{region 'Documentation'}
(*!
<summary>Contributes only the checking Assertions, not the intentionally controlled subject results.</summary>
*)
{endregion}
METHOD PROTECTED AggregateResults
VAR_INPUT
    Aggregator : I_ResultAggregator; //! Borrowed result sink owned by the outer Test Case; add this test's checking Assertions without resetting or retaining the sink.
END_VAR
Aggregator.AddProvider(Provider := FInitialization);
Aggregator.AddProvider(Provider := FConfigureOrder);
Aggregator.AddProvider(Provider := FCollection);
Aggregator.AddProvider(Provider := FPassiveState);
Aggregator.AddProvider(Provider := FDiagnostic);
Aggregator.AddProvider(Provider := FDispatch);
Aggregator.AddProvider(Provider := FCaptureIntegrity);
END_METHOD

{region 'Documentation'}
(*!
<summary>Changes one setup condition and records initialization evidence before cyclic subject execution.</summary>
*)
{endregion}
METHOD PRIVATE BeginAttempt
VAR
    Config : ST_TestSuiteConfig;
    Parent : I_RunControl;
    SuiteName : STRING(GVL_Constants.NameLength);
    Initialized : BOOL;
    ExpectedConfigured : BOOL;
    ExpectedHelper : BOOL;
    Index : UINT;
    FirstChild : I_Orchestratable;
    LastChild : I_Orchestratable;
    SubjectCollection : I_OrchestratableCollection;
    Publisher : I_EventPublisher;
    SubjectStatus : ST_TestSuiteStatus;
    FirstSharedChild : I_Orchestratable;
    LastSharedChild : I_Orchestratable;
    BelowRangeChild : I_Orchestratable;
    UnusedChild : I_Orchestratable;
    UnusedTypedChild : I_TestCase;
END_VAR
FFixtureValid := FCapture.Initialize(Buffer := FEvents,
    FifoControl := FCaptureFifo,
    Status := FCaptureStatus);
IF NOT FFixtureValid THEN
    Error(Message := 'Suite initialization capture could not be initialized.');
    RETURN;
END_IF;
Parent := FSubjectParent;
SuiteName := 'Subject';
CASE FAttempt OF
    MissingParent:
        Parent := 0;
    InvalidName:
        SuiteName := 'Invalid.Subject';
    OverlengthName:
        FOR Index := 1 TO GVL_Constants.NameLength DO
            SuiteName := CONCAT(SuiteName, 'x');
        END_FOR;
    ZeroExecutionTimeout:
        Config.Timeout := T#0s;
    ZeroResetTimeout:
        Config.ResetTimeout := T#0s;
    ZeroAbortTimeout:
        Config.AbortTimeout := T#0s;
ELSE
    // Remaining attempts vary the concrete setup or helper, not these external inputs.
END_CASE;
FExpectedInitialized := (FAttempt = FirstValidSetup) OR (FAttempt = FinalValidSetup);
ExpectedConfigured := FExpectedInitialized OR (FAttempt >= NoRegistration);
ExpectedHelper := ExpectedConfigured AND (FAttempt <> NoRegistration);
FHelper.BeginScenario(AcceptInitialization := FAttempt <> RejectedHelper);
FSubject.Bind(Publisher := FCapture,
    Helper := FHelper,
    RegisterChildren := FAttempt <> NoRegistration,
    IncludeUninitializedChild := FAttempt = UninitializedChild);
Initialized := FSubject.Initialize(Parent := Parent,
    SuiteName := SuiteName,
    ResourceName := 'Fixture',
    Config := Config);
Publisher := FCapture;
SubjectStatus := FSubject.Status;
FInitializationMatches := (Initialized = FExpectedInitialized)
    AND (FSubject.IsInitialized = FExpectedInitialized)
    AND (SubjectStatus.Execution.ConfigError <> FExpectedInitialized)
    AND (FSubject.EventPublisher = Publisher);
FConfigureOrderMatches := FSubject.ConfigureCount = BOOL_TO_UINT(ExpectedConfigured);
IF ExpectedConfigured THEN
    FConfigureOrderMatches := FConfigureOrderMatches AND FSubject.ConfigureContextValid;
END_IF;
FCollectionMatches := FHelper.InitializeCount = BOOL_TO_UINT(ExpectedHelper);
IF ExpectedHelper THEN
    SubjectCollection := FSubject;
    FCollectionMatches := FCollectionMatches
        AND (FHelper.Collection = SubjectCollection)
        AND (FHelper.FirstIndex = 4) AND (FHelper.LastIndex = 6) AND (FHelper.ChildCount = 2)
        AND (FHelper.FirstChild <> 0) AND (FHelper.LastChild <> 0)
        AND (FHelper.FirstChild <> FHelper.LastChild)
        AND (FHelper.OwnerName = FSubject.Name) AND (FHelper.ResourceName = 'Fixture');
END_IF;
FirstSharedChild := FSubject.GetChild(Index := 4);
LastSharedChild := FSubject.GetChild(Index := 5);
BelowRangeChild := FSubject.GetChild(Index := 3);
UnusedChild := FSubject.GetChild(Index := 6);
UnusedTypedChild := FSubject.GetTestCase(Index := 6);
IF FExpectedInitialized THEN
    FirstChild := FSubject.GetTestCase(Index := 4);
    LastChild := FSubject.GetTestCase(Index := 5);
    FCollectionMatches := FCollectionMatches
        AND (FSubject.ChildCount = 2)
        AND (FSubject.ChildArrayLowerBound = 4) AND (FSubject.ChildArrayUpperBound = 6)
        AND (FirstSharedChild = FirstChild)
        AND (LastSharedChild = LastChild)
        AND (FHelper.FirstChild = FirstChild) AND (FHelper.LastChild = LastChild)
        AND (BelowRangeChild = 0) AND (UnusedChild = 0)
        AND (UnusedTypedChild = 0)
        AND (FSubject.Name = CONCAT(FSubjectParent.Name, '.Subject'));
ELSE
    FirstChild := FSubject.GetTestCase(Index := 4);
    FCollectionMatches := FCollectionMatches
        AND (FSubject.ChildCount = 0)
        AND (FSubject.ChildArrayLowerBound = 0) AND (FSubject.ChildArrayUpperBound = 0)
        AND (FirstSharedChild = 0) AND (FirstChild = 0);
END_IF;
FInitialSequence := FCaptureStatus.SequenceId;
IF FExpectedInitialized THEN
    FDiagnosticMatches := FInitialSequence = 0;
ELSE
    FDiagnosticMatches := (FInitialSequence = 1)
        AND (FEvents[1].EventType = E_EventType.Framework)
        AND (FEvents[1].Severity = E_EventSeverity.Error)
        AND (FEvents[1].State = E_State.Uninitialized)
        AND (FEvents[1].Name = FSubject.Name);
END_IF;
FPassiveStateMatches := (FSubject.State = E_State.Uninitialized) AND NOT FSubject.IsReady;
FDispatchMatches := (FHelper.ExecuteCount = 0) AND (FSubject.ChildCallCount = 0);
FPassiveCalls := 0;
FAttemptStarted := TRUE;
END_METHOD

{region 'Documentation'}
(*!
<summary>Supplies only the root identity; the root never executes this isolated subject.</summary>
*)
{endregion}
METHOD PUBLIC BindSubjectParent
VAR_INPUT
    Parent : I_RunControl; //! Borrowed identity parent retained for isolated subject initialization; keep the Run-Control alive through subject use.
END_VAR
FSubjectParent := Parent;
END_METHOD

{region 'Documentation'}
(*!
<summary>Initializes the checking Assertions; the scenario explicitly initializes its isolated subject.</summary>
*)
{endregion}
METHOD PROTECTED Configure
FPreparationStateCount := 0;
FTestStateCount := AttemptCount;
FInitialization.Initialize(Parent := THIS^,
    AssertionName := 'Initialization');
FConfigureOrder.Initialize(Parent := THIS^,
    AssertionName := 'ConfigureOrder');
FCollection.Initialize(Parent := THIS^,
    AssertionName := 'Collection');
FPassiveState.Initialize(Parent := THIS^,
    AssertionName := 'PassiveState');
FDiagnostic.Initialize(Parent := THIS^,
    AssertionName := 'Diagnostic');
FDispatch.Initialize(Parent := THIS^,
    AssertionName := 'Dispatch');
FCaptureIntegrity.Initialize(Parent := THIS^,
    AssertionName := 'CaptureIntegrity');
END_METHOD

{region 'Documentation'}
(*!
<summary>No asynchronous test resource remains to stop.</summary>
*)
{endregion}
METHOD PROTECTED ProcessAbort
VAR_INPUT
    Enable : BOOL; //! Phase permission supplied by the owning Test Case; FALSE does not authorize progression, while observation may continue.
END_VAR
IF Enable THEN
    CompleteAbort();
END_IF;
END_METHOD

{region 'Documentation'}
(*!
<summary>Latches each setup attempt after two passive calls; no automatic Reset or repeated diagnostics are permitted.</summary>
*)
{endregion}
METHOD PROTECTED ProcessAssertions
VAR_INPUT
    Enable : BOOL; //! Phase permission supplied by the owning Test Case; FALSE does not authorize progression, while observation may continue.
END_VAR
VAR
    Evaluate : BOOL;
END_VAR
Evaluate := Enable AND (FPassiveCalls >= PassiveCallCount);
FInitialization(Enable := Evaluate,
    State := State,
    IN := FInitializationMatches);
FConfigureOrder(Enable := Evaluate,
    State := State,
    IN := FConfigureOrderMatches);
FCollection(Enable := Evaluate,
    State := State,
    IN := FCollectionMatches);
FPassiveState(Enable := Evaluate,
    State := State,
    IN := FPassiveStateMatches);
FDiagnostic(Enable := Evaluate,
    State := State,
    IN := FDiagnosticMatches);
FDispatch(Enable := Evaluate,
    State := State,
    IN := FDispatchMatches);
FCaptureIntegrity(Enable := Evaluate,
    State := State,
    IN := FCaptureStatus.LostEventCount = 0);
IF Evaluate THEN
    FChecked := TRUE;
END_IF;
END_METHOD

{region 'Documentation'}
(*!
<summary>No resource Preparation is required for this controlled owner scenario.</summary>
*)
{endregion}
METHOD PROTECTED ProcessPreparations
VAR_INPUT
    // SA0033: Required override; the scenario has no Preparation phase.
    {attribute 'analysis' := '-33'}
    Enable : BOOL; //! Phase permission supplied by the owning Test Case; FALSE does not authorize progression, while observation may continue.
END_VAR
END_METHOD

{region 'Documentation'}
(*!
<summary>Restarts the test script and clears checking Assertions; subject setup belongs to the next test attempt.</summary>
*)
{endregion}
METHOD PROTECTED ProcessReset
FAttempt := FirstValidSetup;
FAttemptStarted := FALSE;
FChecked := FALSE;
FPassiveCalls := 0;
FInitialization.Reset();
FConfigureOrder.Reset();
FCollection.Reset();
FPassiveState.Reset();
FDiagnostic.Reset();
FDispatch.Reset();
FCaptureIntegrity.Reset();
CompleteReset();
END_METHOD

{region 'Documentation'}
(*!
<summary>Advances the explicit test script with at most one subject FB call per active PLC cycle.</summary>
*)
{endregion}
METHOD PROTECTED ProcessTests
VAR_INPUT
    Enable : BOOL; //! Phase permission supplied by the owning Test Case; FALSE does not authorize progression, while observation may continue.
END_VAR
IF NOT Enable THEN
    RETURN;
END_IF;
IF FChecked THEN
    IF FAttempt = AttemptCount THEN
        CompleteTests();
        RETURN;
    END_IF;
    FAttempt := FAttempt + 1;
    FAttemptStarted := FALSE;
    FChecked := FALSE;
    NextTestState();
END_IF;
IF NOT FAttemptStarted THEN
    BeginAttempt();
    IF NOT FFixtureValid THEN
        RETURN;
    END_IF;
END_IF;
FSubject();
FPassiveCalls := FPassiveCalls + 1;
FPassiveStateMatches := FPassiveStateMatches
    AND (FSubject.State = E_State.Uninitialized)
    AND NOT FSubject.IsReady
    AND (FSubject.Result = E_Result.NotEvaluated);
IF FExpectedInitialized THEN
    FDispatchMatches := FDispatchMatches
        AND (FHelper.ExecuteCount = FPassiveCalls)
        AND (FSubject.ChildCallCount = FPassiveCalls)
        AND (FHelper.CurrentTask = E_OrchestratorTask.Idle);
ELSE
    FDispatchMatches := FDispatchMatches
        AND (FHelper.ExecuteCount = 0) AND (FSubject.ChildCallCount = 0);
END_IF;
FDiagnosticMatches := FDiagnosticMatches AND (FCaptureStatus.SequenceId = FInitialSequence);
END_METHOD

END_FUNCTION_BLOCK

// ---- SelfTests/TestCases/TestSuite_TestSuiteLifecycle/Helper/TestSuiteLifecycleProbe.TcPOU
{region 'Documentation'}
(*!
<summary>Thin TestSuiteBase subject with a typed child array and isolated dependencies.</summary>
<description>
Bind is called before Initialize. Production initialization, sequencing, aggregation and
publication remain inherited. Configure records its context and builds a small real collection.
The uninitialized-child option uses a separate never-initialized double, not mutated base state.
ProcessTestCases applies the scenario's child view only after the base has called its helper.
</description>
*)
{endregion}
FUNCTION_BLOCK TestSuiteLifecycleProbe EXTENDS TestSuiteBase
VAR
    FChildA : SuiteLifecycleChildDouble;
    FChildB : SuiteLifecycleChildDouble;
    FUninitializedChild : SuiteLifecycleChildDouble;
    FTestCases : ARRAY[4..6] OF I_TestCase;
    FChildObservation : ST_OrchestrationObservation;
    FSecondChildObservation : ST_OrchestrationObservation;
    FRegisterChildren : BOOL := TRUE;
    FIncludeUninitializedChild : BOOL;
    FConfigureCount : UINT;
    FConfigureContextValid : BOOL;
    FChildCallCount : UINT;
END_VAR

SUPER^();

{region 'Documentation'}
(*!
<summary>Binds isolated dependencies before Initialize and selects the concrete setup to exercise.</summary>
*)
{endregion}
METHOD PUBLIC Bind
VAR_INPUT
    Publisher : I_EventPublisher; //! Nonzero isolated event publisher retained before subject initialization; keep it alive through all subject use.
    Helper : I_Orchestrator; //! Nonzero injected orchestration helper retained before owner initialization; keep it alive through subject use.
    RegisterChildren : BOOL := TRUE; //! TRUE registers the two controlled children; FALSE exercises empty configuration.
    IncludeUninitializedChild : BOOL := FALSE; //! TRUE leaves a registered controlled child uninitialized to exercise rejection.
END_VAR
FEventPublisher := Publisher;
FOrchestrator := Helper;
FRegisterChildren := RegisterChildren;
FIncludeUninitializedChild := IncludeUninitializedChild;
FChildA.SetReleaseResponse();
FChildB.SetReleaseResponse();
FConfigureCount := 0;
FChildCallCount := 0;
FConfigureContextValid := FALSE;
FChildObservation.State := E_State.Uninitialized;
FChildObservation.Result := E_Result.NotEvaluated;
FChildObservation.Ready := FALSE;
FChildObservation.Complete := FALSE;
FSecondChildObservation := FChildObservation;
END_METHOD

{region 'Documentation'}
(*!
<summary>Both concrete child bodies have executed exactly once per ProcessTestCases invocation.</summary>
*)
{endregion}
{attribute 'monitoring' := 'call'}
PROPERTY PUBLIC ChildBodyCallsMatch : BOOL //! Both concrete child bodies have executed exactly once per ProcessTestCases invocation.
GET
VAR
    FirstCalls : ST_OrchestrationCalls;
    SecondCalls : ST_OrchestrationCalls;
END_VAR
FirstCalls := FChildA.Calls;
SecondCalls := FChildB.Calls;
ChildBodyCallsMatch := (FirstCalls.BodyCount = FChildCallCount) AND (SecondCalls.BodyCount = FChildCallCount);
END_GET
END_PROPERTY

{region 'Documentation'}
(*!
<summary>Number of ProcessTestCases invocations since binding.</summary>
*)
{endregion}
{attribute 'monitoring' := 'call'}
PROPERTY PUBLIC ChildCallCount : UINT //! Number of ProcessTestCases invocations since binding.
GET
ChildCallCount := FChildCallCount;
END_GET
END_PROPERTY

{region 'Documentation'}
(*!
<summary>Registers two controlled typed children in a shifted array with spare capacity; records base context.</summary>
*)
{endregion}
METHOD PROTECTED Configure
VAR_IN_OUT
    // SA0167: Borrowed setup builder; no temporary instance is created.
    {attribute 'analysis' := '-167'}
    Builder : TestSuiteConfigurationBuilder; //! Borrowed owner configuration builder used only during this Configure call; register this owner's concrete children.
END_VAR
FConfigureCount := FConfigureCount + 1;
FConfigureContextValid := (State = E_State.Uninitialized) AND NOT IsInitialized AND (Name <> '');
Builder.Initialize(Mode := E_OrchestrationMode.Serial,
    TestCases := FTestCases);
FChildA.Initialize(Name := CONCAT(Name, '.ChildA'),
    Slot := 0);
FChildB.Initialize(Name := CONCAT(Name, '.ChildB'),
    Slot := 0);
IF NOT FRegisterChildren THEN
    RETURN;
END_IF;
Builder.Register(TestCase := FChildA);
IF FIncludeUninitializedChild THEN
    Builder.Register(TestCase := FUninitializedChild);
ELSE
    Builder.Register(TestCase := FChildB);
END_IF;
END_METHOD

{region 'Documentation'}
(*!
<summary>Configure saw the new identity before successful initialization.</summary>
*)
{endregion}
{attribute 'monitoring' := 'call'}
PROPERTY PUBLIC ConfigureContextValid : BOOL //! Configure saw the new identity before successful initialization.
GET
ConfigureContextValid := FConfigureContextValid;
END_GET
END_PROPERTY

{region 'Documentation'}
(*!
<summary>Number of Configure calls since binding.</summary>
*)
{endregion}
{attribute 'monitoring' := 'call'}
PROPERTY PUBLIC ConfigureCount : UINT //! Number of Configure calls since binding.
GET
ConfigureCount := FConfigureCount;
END_GET
END_PROPERTY

{region 'Documentation'}
(*!
<summary>Returns the recorded calls of a registered controlled child; unknown indices return an empty observation.</summary>
*)
{endregion}
METHOD PUBLIC GetChildCalls : ST_OrchestrationCalls //! Retained call trace for the selected child; an empty trace for an unknown index or empty collection.
VAR_INPUT
    Index : DINT; //! Original occupied child-array index; unknown indices return an empty trace.
END_VAR
VAR
    EmptyCalls : ST_OrchestrationCalls;
END_VAR
GetChildCalls := EmptyCalls;
IF ChildCount = 0 THEN
    RETURN;
END_IF;
IF Index = ChildArrayLowerBound THEN
    GetChildCalls := FChildA.Calls;
ELSIF (ChildCount > 1) AND (Index = ChildArrayLowerBound + 1) THEN
    GetChildCalls := FChildB.Calls;
END_IF;
END_METHOD

{region 'Documentation'}
(*!
<summary>Returns the registered typed entry by actual array index; lookup never executes a child.</summary>
*)
{endregion}
METHOD PUBLIC GetTestCase : I_TestCase //! Typed child interface at the original array index; zero when no entry is available.
VAR_INPUT
    Index : DINT; //! Original occupied child-array index, rather than an ordinal position.
END_VAR
GetTestCase := 0;
IF (ChildCount = 0) OR (Index < ChildArrayLowerBound)
    OR (DINT_TO_LINT(Index) >= DINT_TO_LINT(ChildArrayLowerBound) + UINT_TO_LINT(ChildCount)) THEN
    RETURN;
END_IF;
GetTestCase := FTestCases[Index];
END_METHOD

{region 'Documentation'}
(*!
<summary>Applies the next scripted observation after the helper; counts calls without replacing owner processing.</summary>
*)
{endregion}
METHOD PROTECTED ProcessTestCases
FChildA(ObservationInput := FChildObservation);
FChildB(ObservationInput := FSecondChildObservation);
FChildCallCount := FChildCallCount + 1;
END_METHOD

{region 'Documentation'}
(*!
<summary>Selects the next child snapshot; it becomes visible only in ProcessTestCases, after helper execution.</summary>
*)
{endregion}
METHOD PUBLIC SetChildObservation
VAR_INPUT
    Observation : ST_OrchestrationObservation; //! Scripted view copied to both children for acceptance on their next concrete body calls.
END_VAR
FChildObservation := Observation;
FSecondChildObservation := Observation;
END_METHOD

{region 'Documentation'}
(*!
<summary>Supplies independent next snapshots; each child accepts its view only when the Suite calls its body.</summary>
*)
{endregion}
METHOD PUBLIC SetChildObservations
VAR_INPUT
    FirstChild : ST_OrchestrationObservation; //! Scripted view for the first child, accepted on its next concrete body call.
    SecondChild : ST_OrchestrationObservation; //! Scripted view for the second child, accepted on its next concrete body call.
END_VAR
FChildObservation := FirstChild;
FSecondChildObservation := SecondChild;
END_METHOD

{region 'Documentation'}
(*!
<summary>Controls only the child release boundary for delegation tests, without changing Suite accounting.</summary>
*)
{endregion}
METHOD PUBLIC SetChildReleaseResponses
VAR_INPUT
    FirstSucceeds : BOOL := TRUE; //! Release response installed in the first controlled child.
    SecondSucceeds : BOOL := TRUE; //! Release response installed in the second controlled child.
END_VAR
FChildA.SetReleaseResponse(Succeeds := FirstSucceeds);
FChildB.SetReleaseResponse(Succeeds := SecondSucceeds);
END_METHOD

END_FUNCTION_BLOCK

// ---- SelfTests/TestCases/TestSuite_TestSuiteLifecycle/Helper/SuiteLifecycleChildDouble.TcPOU
{region 'Documentation'}
(*!
<summary>Adds the typed Test Case status to the existing scripted child boundary; requests remain observation-only.</summary>
*)
{endregion}
FUNCTION_BLOCK SuiteLifecycleChildDouble EXTENDS OrchestrationChildDouble IMPLEMENTS I_TestCase
VAR
    FReleaseSucceeds : BOOL := TRUE;
END_VAR

SUPER^(ObservationInput := ObservationInput);

{region 'Documentation'}
(*!
<summary>Records a scripted rejection without release; successful calls use the original double's release behavior.</summary>
*)
{endregion}
METHOD PUBLIC FreeReservedEvents : BOOL //! FALSE for scripted rejection; otherwise the original double release result.
IF NOT FReleaseSucceeds THEN
    FCalls.FreeCount := FCalls.FreeCount + 1;
    FreeReservedEvents := FALSE;
    RETURN;
END_IF;
FreeReservedEvents := SUPER^.FreeReservedEvents();
END_METHOD

{region 'Documentation'}
(*!
<summary>Controls release success without altering the marker or call observations.</summary>
*)
{endregion}
METHOD PUBLIC SetReleaseResponse
VAR_INPUT
    Succeeds : BOOL := TRUE; //! FALSE scripts release rejection without clearing the local marker; TRUE delegates normal release.
END_VAR
FReleaseSucceeds := Succeeds;
END_METHOD

{region 'Documentation'}
(*!
<summary>Projects the scripted child observation into the typed Suite-facing status; no lifecycle is copied.</summary>
*)
{endregion}
{attribute 'monitoring' := 'variable'}
PROPERTY PUBLIC Status : ST_TestCaseStatus //! Projects the scripted child observation into the typed Suite-facing status; no lifecycle is copied.
GET
VAR
    Snapshot : ST_TestCaseStatus;
    View : ST_OrchestrationObservation;
END_VAR
View := Observation;
Snapshot.Execution.State := View.State;
Snapshot.Execution.Result := View.Result;
Snapshot.Execution.Ready := View.Ready;
Snapshot.Execution.Completed := View.Complete;
Snapshot.Execution.Error := View.Result = E_Result.Error;
CASE View.State OF
    E_State.Uninitialized:
        Snapshot.Execution.ExecutionStatus := E_ExecutionStatus.NotReady;
        Snapshot.Execution.Uninitialized := TRUE;
    E_State.Reset:
        Snapshot.Execution.ExecutionStatus := E_ExecutionStatus.Reset;
    E_State.Idle:
        Snapshot.Execution.ExecutionStatus := E_ExecutionStatus.Idle;
    E_State.Starting:
        Snapshot.Execution.ExecutionStatus := E_ExecutionStatus.Starting;
    E_State.Running:
        Snapshot.Execution.ExecutionStatus := E_ExecutionStatus.Running;
        Snapshot.Execution.Running := TRUE;
    E_State.Completing:
        Snapshot.Execution.ExecutionStatus := E_ExecutionStatus.Completing;
    E_State.Completed:
        Snapshot.Execution.ExecutionStatus := E_ExecutionStatus.Completed;
    E_State.Aborting, E_State.AbortingFromError:
        Snapshot.Execution.ExecutionStatus := E_ExecutionStatus.Aborting;
ELSE
    Snapshot.Execution.ExecutionStatus := E_ExecutionStatus.Error;
END_CASE;
Status := Snapshot;
END_GET
END_PROPERTY

END_FUNCTION_BLOCK

// ---- SelfTests/TestCases/TestSuite_TestSuiteLifecycle/Helper/SuiteOrchestratorDouble.TcPOU
{region 'Documentation'}
(*!
<summary>Controlled I_Orchestrator boundary for Suite owner tests, without a scheduler.</summary>
<description>
Initialize records identity, collection bounds and child identities while the owner is still
initializing. Execute records task assignment and pre-child-call states. SetObservation supplies deliberate
responses between owner cycles; no child requests, reservations or state machine are copied.
The test supplies coherent child observations separately through the concrete Suite adapter.
</description>
*)
{endregion}
FUNCTION_BLOCK SuiteOrchestratorDouble IMPLEMENTS I_Orchestrator
VAR
    FAcceptInitialization : BOOL := TRUE;
    FInitialized : BOOL;
    FInitializeCount : UINT;
    FExecuteCount : UINT;
    FFirstChildStateAtExecute : E_State;
    FLastChildStateAtExecute : E_State;
    FCurrentTask : E_OrchestratorTask;
    FCollection : I_OrchestratableCollection;
    FName : STRING(GVL_Constants.NameLength);
    FResourceName : STRING(GVL_Constants.ResourceNameLength);
    FFirstIndex : DINT;
    FLastIndex : DINT;
    FChildCount : UINT;
    FFirstChild : I_Orchestratable;
    FLastChild : I_Orchestratable;
    FReady : BOOL;
    FResult : E_Result;
    FResetFinished : BOOL;
    FAbortFinished : BOOL;
    FExecutionFinished : BOOL;
END_VAR

{region 'Documentation'}
(*!
<summary>Clears observations before owner initialization and selects only the initialization outcome.</summary>
*)
{endregion}
METHOD PUBLIC BeginScenario
VAR_INPUT
    AcceptInitialization : BOOL := TRUE; //! Scripted acceptance returned by subsequent Initialize calls.
END_VAR
FAcceptInitialization := AcceptInitialization;
FInitialized := FALSE;
FInitializeCount := 0;
FExecuteCount := 0;
FFirstChildStateAtExecute := E_State.Uninitialized;
FLastChildStateAtExecute := E_State.Uninitialized;
FCurrentTask := E_OrchestratorTask.Idle;
FCollection := 0;
FName := '';
FResourceName := '';
FFirstIndex := 0;
FLastIndex := 0;
FChildCount := 0;
FFirstChild := 0;
FLastChild := 0;
SetObservation(Ready := FALSE);
END_METHOD

{region 'Documentation'}
(*!
<summary>Population observed synchronously inside Initialize.</summary>
*)
{endregion}
{attribute 'monitoring' := 'call'}
PROPERTY PUBLIC ChildCount : UINT //! Population observed synchronously inside Initialize.
GET
ChildCount := FChildCount;
END_GET
END_PROPERTY

{region 'Documentation'}
(*!
<summary>The exact collection interface supplied by the owner.</summary>
*)
{endregion}
{attribute 'monitoring' := 'variable'}
PROPERTY PUBLIC Collection : I_OrchestratableCollection //! The exact collection interface supplied by the owner.
GET
Collection := FCollection;
END_GET
END_PROPERTY

{region 'Documentation'}
(*!
<summary>Last task supplied by the owner.</summary>
*)
{endregion}
{attribute 'monitoring' := 'call'}
PROPERTY PUBLIC CurrentTask : E_OrchestratorTask //! Last task supplied by the owner.
GET
CurrentTask := FCurrentTask;
END_GET
END_PROPERTY

{region 'Documentation'}
(*!
<summary>Records the owner task and current child states; no observations are changed or child commands sent.</summary>
*)
{endregion}
METHOD PUBLIC Execute
VAR_INPUT
    Task : E_OrchestratorTask; //! Owner-assigned task to record; this double does not execute or request children.
END_VAR
FCurrentTask := Task;
FExecuteCount := FExecuteCount + 1;
IF FFirstChild <> 0 THEN
    FFirstChildStateAtExecute := FFirstChild.State;
END_IF;
IF FLastChild <> 0 THEN
    FLastChildStateAtExecute := FLastChild.State;
END_IF;
END_METHOD

{region 'Documentation'}
(*!
<summary>Number of cyclic helper calls.</summary>
*)
{endregion}
{attribute 'monitoring' := 'call'}
PROPERTY PUBLIC ExecuteCount : UINT //! Number of cyclic helper calls.
GET
ExecuteCount := FExecuteCount;
END_GET
END_PROPERTY

{region 'Documentation'}
(*!
<summary>First occupied interface observed inside Initialize.</summary>
*)
{endregion}
{attribute 'monitoring' := 'variable'}
PROPERTY PUBLIC FirstChild : I_Orchestratable //! First occupied interface observed inside Initialize.
GET
FirstChild := FFirstChild;
END_GET
END_PROPERTY

{region 'Documentation'}
(*!
<summary>First child state observed by the helper before concrete child calls.</summary>
*)
{endregion}
{attribute 'monitoring' := 'call'}
PROPERTY PUBLIC FirstChildStateAtExecute : E_State //! First child state observed by the helper before concrete child calls.
GET
FirstChildStateAtExecute := FFirstChildStateAtExecute;
END_GET
END_PROPERTY

{region 'Documentation'}
(*!
<summary>Lower bound observed synchronously inside Initialize.</summary>
*)
{endregion}
{attribute 'monitoring' := 'call'}
PROPERTY PUBLIC FirstIndex : DINT //! Lower bound observed synchronously inside Initialize.
GET
FirstIndex := FFirstIndex;
END_GET
END_PROPERTY

{region 'Documentation'}
(*!
<summary>Records and immediately queries the collection handed over by the owner; never executes children.</summary>
*)
{endregion}
METHOD PUBLIC Initialize : BOOL //! Scripted initialization acceptance; the supplied collection is queried regardless of that response.
VAR_INPUT
    Collection : I_OrchestratableCollection; //! Nonzero borrowed collection queried immediately and retained; keep the collection and children alive.
    Name : STRING(GVL_Constants.NameLength); //! Owner diagnostic name retained by the double.
    ResourceName : STRING(GVL_Constants.ResourceNameLength) := ''; //! Owner diagnostic resource retained by the double.
END_VAR
FInitializeCount := FInitializeCount + 1;
FCollection := Collection;
FName := Name;
FResourceName := ResourceName;
FFirstIndex := Collection.ChildArrayLowerBound;
FLastIndex := Collection.ChildArrayUpperBound;
FChildCount := Collection.ChildCount;
IF FChildCount > 0 THEN
    FFirstChild := Collection.GetChild(Index := FFirstIndex);
    FLastChild := Collection.GetChild(Index := FFirstIndex + UINT_TO_DINT(FChildCount) - 1);
END_IF;
FInitialized := FAcceptInitialization;
Initialize := FInitialized;
END_METHOD

{region 'Documentation'}
(*!
<summary>Number of owner initialization calls.</summary>
*)
{endregion}
{attribute 'monitoring' := 'call'}
PROPERTY PUBLIC InitializeCount : UINT //! Number of owner initialization calls.
GET
InitializeCount := FInitializeCount;
END_GET
END_PROPERTY

{region 'Documentation'}
(*!
<summary>Scripted Abort completion.</summary>
*)
{endregion}
{attribute 'monitoring' := 'call'}
PROPERTY PUBLIC IsAbortFinished : BOOL //! Scripted Abort completion.
GET
IsAbortFinished := FAbortFinished;
END_GET
END_PROPERTY

{region 'Documentation'}
(*!
<summary>Scripted execution completion.</summary>
*)
{endregion}
{attribute 'monitoring' := 'call'}
PROPERTY PUBLIC IsExecutionFinished : BOOL //! Scripted execution completion.
GET
IsExecutionFinished := FExecutionFinished;
END_GET
END_PROPERTY

{region 'Documentation'}
(*!
<summary>Accepted initialization response.</summary>
*)
{endregion}
{attribute 'monitoring' := 'call'}
PROPERTY PUBLIC IsInitialized : BOOL //! Accepted initialization response.
GET
IsInitialized := FInitialized;
END_GET
END_PROPERTY

{region 'Documentation'}
(*!
<summary>Scripted child readiness summary.</summary>
*)
{endregion}
{attribute 'monitoring' := 'call'}
PROPERTY PUBLIC IsReady : BOOL //! Scripted child readiness summary.
GET
IsReady := FReady;
END_GET
END_PROPERTY

{region 'Documentation'}
(*!
<summary>Whether the owner currently assigns Reset.</summary>
*)
{endregion}
{attribute 'monitoring' := 'call'}
PROPERTY PUBLIC IsResetActive : BOOL //! Whether the owner currently assigns Reset.
GET
IsResetActive := FCurrentTask = E_OrchestratorTask.Reset;
END_GET
END_PROPERTY

{region 'Documentation'}
(*!
<summary>Scripted Reset completion.</summary>
*)
{endregion}
{attribute 'monitoring' := 'call'}
PROPERTY PUBLIC IsResetFinished : BOOL //! Scripted Reset completion.
GET
IsResetFinished := FResetFinished;
END_GET
END_PROPERTY

{region 'Documentation'}
(*!
<summary>Last occupied interface observed inside Initialize.</summary>
*)
{endregion}
{attribute 'monitoring' := 'variable'}
PROPERTY PUBLIC LastChild : I_Orchestratable //! Last occupied interface observed inside Initialize.
GET
LastChild := FLastChild;
END_GET
END_PROPERTY

{region 'Documentation'}
(*!
<summary>Last child state observed by the helper before concrete child calls.</summary>
*)
{endregion}
{attribute 'monitoring' := 'call'}
PROPERTY PUBLIC LastChildStateAtExecute : E_State //! Last child state observed by the helper before concrete child calls.
GET
LastChildStateAtExecute := FLastChildStateAtExecute;
END_GET
END_PROPERTY

{region 'Documentation'}
(*!
<summary>Capacity upper bound observed synchronously inside Initialize.</summary>
*)
{endregion}
{attribute 'monitoring' := 'call'}
PROPERTY PUBLIC LastIndex : DINT //! Capacity upper bound observed synchronously inside Initialize.
GET
LastIndex := FLastIndex;
END_GET
END_PROPERTY

{region 'Documentation'}
(*!
<summary>Diagnostic identity supplied by the owner.</summary>
*)
{endregion}
{attribute 'monitoring' := 'variable'}
PROPERTY PUBLIC OwnerName : STRING(GVL_Constants.NameLength) //! Diagnostic identity supplied by the owner.
GET
OwnerName := FName;
END_GET
END_PROPERTY

{region 'Documentation'}
(*!
<summary>Diagnostic resource supplied by the owner.</summary>
*)
{endregion}
{attribute 'monitoring' := 'variable'}
PROPERTY PUBLIC ResourceName : STRING(GVL_Constants.ResourceNameLength) //! Diagnostic resource supplied by the owner.
GET
ResourceName := FResourceName;
END_GET
END_PROPERTY

{region 'Documentation'}
(*!
<summary>Scripted helper technical result.</summary>
*)
{endregion}
{attribute 'monitoring' := 'call'}
PROPERTY PUBLIC Result : E_Result //! Scripted helper technical result.
GET
Result := FResult;
END_GET
END_PROPERTY

{region 'Documentation'}
(*!
<summary>Supplies the interface response for the next owner call; defaults describe unfinished neutral work.</summary>
*)
{endregion}
METHOD PUBLIC SetObservation
VAR_INPUT
    Ready : BOOL; //! Scripted readiness returned to the owner.
    Result : E_Result := E_Result.NotEvaluated; //! Scripted helper technical result returned to the owner.
    ResetFinished : BOOL := FALSE; //! Scripted Reset-completion signal returned to the owner.
    AbortFinished : BOOL := FALSE; //! Scripted Abort-completion signal returned to the owner.
    ExecutionFinished : BOOL := FALSE; //! Scripted execution-completion signal returned to the owner.
END_VAR
FReady := Ready;
FResult := Result;
FResetFinished := ResetFinished;
FAbortFinished := AbortFinished;
FExecutionFinished := ExecutionFinished;
END_METHOD

END_FUNCTION_BLOCK

// ---- SelfTests/TestCases/TestSuite_TestSuiteLifecycle/Test_SuiteReadiness.TcPOU
{region 'Documentation'}
(*!
<summary>Checks that Suite Start is authorized by owner state and the selected helper's readiness and result.</summary>
<description>
The real Suite reaches Idle through its normal Reset path. The helper then withholds readiness
while the child snapshots are already ready, as can occur before cleanup is observed.
A denied Start must not remain queued when readiness later arrives. A subsequent helper Error
must prevent Start and propagate to the Suite, without selecting helper Execution.
No child scheduling is simulated: controlled snapshots and helper responses isolate owner decisions.
</description>
*)
{endregion}
FUNCTION_BLOCK Test_SuiteReadiness EXTENDS TestCaseBase
VAR
    FSubjectParent : I_RunControl;
    FSubject : TestSuiteLifecycleProbe;
    FHelper : SuiteOrchestratorDouble;
    FCapture : EventBuffer;
    FEvents : ARRAY[1..CaptureLength] OF ST_Event;
    FCaptureFifo : ST_FifoStatus;
    FCaptureStatus : ST_EventBufferStatus;
    FStep : INT;
    FChecked : BOOL;
    FInitialization : AssertTrue;
    FInitializationMatches : BOOL := TRUE;
    FReadiness : AssertTrue;
    FReadinessMatches : BOOL := TRUE;
    FStartGate : AssertTrue;
    FStartGateMatches : BOOL := TRUE;
    FHelperBinding : AssertTrue;
    FHelperBindingMatches : BOOL := TRUE;
    FCaptureIntegrity : AssertTrue;
    FCaptureIntegrityMatches : BOOL := TRUE;
END_VAR
VAR CONSTANT
    CaptureLength : UINT := 64;
    Setup : INT := 0;
    ResetRequested : INT := 1;
    ResetCompleted : INT := 2;
    DenyStart : INT := 3;
    ReleaseReadiness : INT := 4;
    RejectHelperError : INT := 5;
    Finished : INT := 6;
END_VAR

SUPER^();

{region 'Documentation'}
(*!
<summary>Contributes only the checking Assertions, not the intentionally controlled subject results.</summary>
*)
{endregion}
METHOD PROTECTED AggregateResults
VAR_INPUT
    Aggregator : I_ResultAggregator; //! Borrowed result sink owned by the outer Test Case; add this test's checking Assertions without resetting or retaining the sink.
END_VAR
Aggregator.AddProvider(Provider := FInitialization);
Aggregator.AddProvider(Provider := FReadiness);
Aggregator.AddProvider(Provider := FStartGate);
Aggregator.AddProvider(Provider := FHelperBinding);
Aggregator.AddProvider(Provider := FCaptureIntegrity);
END_METHOD

{region 'Documentation'}
(*!
<summary>Supplies only the root identity; the root never executes this isolated subject.</summary>
*)
{endregion}
METHOD PUBLIC BindSubjectParent
VAR_INPUT
    Parent : I_RunControl; //! Borrowed identity parent retained for isolated subject initialization; keep the Run-Control alive through subject use.
END_VAR
FSubjectParent := Parent;
END_METHOD

{region 'Documentation'}
(*!
<summary>Initializes the checking Assertions; the scenario explicitly initializes its isolated subject.</summary>
*)
{endregion}
METHOD PROTECTED Configure
FPreparationStateCount := 0;
FTestStateCount := 1;
FInitialization.Initialize(Parent := THIS^,
    AssertionName := 'Initialization');
FReadiness.Initialize(Parent := THIS^,
    AssertionName := 'Readiness');
FStartGate.Initialize(Parent := THIS^,
    AssertionName := 'StartGate');
FHelperBinding.Initialize(Parent := THIS^,
    AssertionName := 'HelperBinding');
FCaptureIntegrity.Initialize(Parent := THIS^,
    AssertionName := 'CaptureIntegrity');
END_METHOD

{region 'Documentation'}
(*!
<summary>No asynchronous test resource remains to stop.</summary>
*)
{endregion}
METHOD PROTECTED ProcessAbort
VAR_INPUT
    Enable : BOOL; //! Phase permission supplied by the owning Test Case; FALSE does not authorize progression, while observation may continue.
END_VAR
IF Enable THEN
    CompleteAbort();
END_IF;
END_METHOD

{region 'Documentation'}
(*!
<summary>Evaluates the complete readiness script and consumes reset requests on disabled calls.</summary>
*)
{endregion}
METHOD PROTECTED ProcessAssertions
VAR_INPUT
    Enable : BOOL; //! Phase permission supplied by the owning Test Case; FALSE does not authorize progression, while observation may continue.
END_VAR
VAR
    Evaluate : BOOL;
END_VAR
Evaluate := Enable AND (FStep = Finished);
FInitialization(Enable := Evaluate,
    State := State,
    IN := FInitializationMatches);
FReadiness(Enable := Evaluate,
    State := State,
    IN := FReadinessMatches);
FStartGate(Enable := Evaluate,
    State := State,
    IN := FStartGateMatches);
FHelperBinding(Enable := Evaluate,
    State := State,
    IN := FHelperBindingMatches);
FCaptureIntegrity(Enable := Evaluate,
    State := State,
    IN := FCaptureIntegrityMatches);
IF Evaluate THEN
    FChecked := TRUE;
END_IF;
END_METHOD

{region 'Documentation'}
(*!
<summary>No resource Preparation is required for this controlled owner scenario.</summary>
*)
{endregion}
METHOD PROTECTED ProcessPreparations
VAR_INPUT
    // SA0033: Required override; the scenario has no Preparation phase.
    {attribute 'analysis' := '-33'}
    Enable : BOOL; //! Phase permission supplied by the owning Test Case; FALSE does not authorize progression, while observation may continue.
END_VAR
END_METHOD

{region 'Documentation'}
(*!
<summary>Restarts the test script and clears checking Assertions; subject setup belongs to the next test attempt.</summary>
*)
{endregion}
METHOD PROTECTED ProcessReset
FStep := Setup;
FChecked := FALSE;
FInitializationMatches := TRUE;
FReadinessMatches := TRUE;
FStartGateMatches := TRUE;
FHelperBindingMatches := TRUE;
FCaptureIntegrityMatches := TRUE;
FInitialization.Reset();
FReadiness.Reset();
FStartGate.Reset();
FHelperBinding.Reset();
FCaptureIntegrity.Reset();
CompleteReset();
END_METHOD

{region 'Documentation'}
(*!
<summary>Advances the explicit test script with at most one subject FB call per active PLC cycle.</summary>
*)
{endregion}
METHOD PROTECTED ProcessTests
VAR_INPUT
    Enable : BOOL; //! Phase permission supplied by the owning Test Case; FALSE does not authorize progression, while observation may continue.
END_VAR
IF NOT Enable THEN
    RETURN;
END_IF;
IF FChecked THEN
    CompleteTests();
    RETURN;
END_IF;
RunStep();
END_METHOD

{region 'Documentation'}
(*!
<summary>Exercises readiness through normal Reset, denied Start, helper release and a held helper error.</summary>
*)
{endregion}
METHOD PRIVATE RunStep
VAR
    Config : ST_TestSuiteConfig;
    ChildView : ST_OrchestrationObservation;
    Initialized : BOOL;
    ExpectedCalls : UINT;
    SubjectStatus : ST_TestSuiteStatus;
END_VAR
CASE FStep OF
    Setup:
        IF NOT FCapture.Initialize(Buffer := FEvents,
            FifoControl := FCaptureFifo,
            Status := FCaptureStatus) THEN
            Error(Message := 'Suite readiness capture could not be initialized.');
            RETURN;
        END_IF;
        FHelper.BeginScenario();
        FSubject.Bind(Publisher := FCapture,
            Helper := FHelper);
        Initialized := FSubject.Initialize(Parent := FSubjectParent,
            SuiteName := 'ReadinessSubject',
            Config := Config);
        FInitializationMatches := Initialized AND FSubject.IsInitialized AND NOT FSubject.IsReady;
        IF NOT Initialized THEN
            FStep := Finished;
            RETURN;
        END_IF;
        FSubject();
        SubjectStatus := FSubject.Status;
        FReadinessMatches := NOT FSubject.IsReady AND (FSubject.State = E_State.Uninitialized);
    ResetRequested:
        IF FSubject.ReserveResetEvents() <> E_EventReservationResult.Accepted THEN
            Error(Message := 'Suite readiness Reset reservation was rejected.');
            RETURN;
        END_IF;
        ChildView.State := E_State.Reset;
        ChildView.Ready := FALSE;
        FSubject.SetChildObservation(Observation := ChildView);
        FSubject.RequestReset();
        FSubject();
        SubjectStatus := FSubject.Status;
        FReadinessMatches := FReadinessMatches AND NOT FSubject.IsReady
            AND (FSubject.State = E_State.Reset);
    ResetCompleted:
        // Ready children alone do not imply that helper cleanup and readiness are complete.
        FSubject.SetChildObservation(Observation := ChildView);
        FHelper.SetObservation(Ready := FALSE,
            ResetFinished := TRUE);
        FSubject();
        SubjectStatus := FSubject.Status;
        FReadinessMatches := FReadinessMatches AND FSubject.IsIdle AND NOT FSubject.IsReady
            AND NOT SubjectStatus.Execution.Ready;
        IF NOT FSubject.FreeReservedEvents() THEN
            Error(Message := 'Suite readiness Reset reservation could not be released.');
            RETURN;
        END_IF;
    DenyStart:
        FHelper.SetObservation(Ready := FALSE);
        FSubject.RequestStart();
        FSubject();
        SubjectStatus := FSubject.Status;
        FStartGateMatches := FSubject.IsIdle
            AND (FHelper.CurrentTask = E_OrchestratorTask.Idle)
            AND NOT FSubject.IsReady;
    ReleaseReadiness:
        FHelper.SetObservation(Ready := TRUE);
        FSubject();
        SubjectStatus := FSubject.Status;
        FReadinessMatches := FReadinessMatches AND FSubject.IsReady
            AND SubjectStatus.Execution.Ready AND FSubject.IsIdle;
        FStartGateMatches := FStartGateMatches
            AND (FHelper.CurrentTask = E_OrchestratorTask.Idle);
    RejectHelperError:
        FHelper.SetObservation(Ready := FALSE,
            Result := E_Result.Error);
        FReadinessMatches := FReadinessMatches AND NOT FSubject.IsReady;
        FSubject.RequestStart();
        FSubject();
        SubjectStatus := FSubject.Status;
        FStartGateMatches := FStartGateMatches
            AND (FSubject.State = E_State.Completing)
            AND (FSubject.Result = E_Result.Error)
            AND (FHelper.CurrentTask = E_OrchestratorTask.Idle);
ELSE
    Error(Message := 'Unexpected Suite readiness test step.');
    RETURN;
END_CASE;
ExpectedCalls := INT_TO_UINT(FStep + 1);
FHelperBindingMatches := FHelperBindingMatches
    AND (FHelper.InitializeCount = 1)
    AND (FHelper.ExecuteCount = ExpectedCalls)
    AND (FSubject.ChildCallCount = ExpectedCalls);
FCaptureIntegrityMatches := FCaptureIntegrityMatches AND (FCaptureStatus.LostEventCount = 0);
FStep := FStep + 1;
END_METHOD

END_FUNCTION_BLOCK

// ---- SelfTests/TestCases/TestSuite_TestSuiteLifecycle/Test_SuiteNormalLifecycle.TcPOU
{region 'Documentation'}
(*!
<summary>Verifies the normal Suite lifecycle with all-Passed or mixed Passed/Failed child results.</summary>
<description>

One owner call per step

Each outer Test state arranges child snapshots and a helper response, calls the real Suite
once, and checks its state, helper task, result and counters. Assertions run before advancing.
The same script is instantiated twice; FirstChildResult stays Passed or Failed for the run.
Both send another Reset while waiting and when the helper finishes; these requests must not
suppress the transition to Idle or change the retained NotEvaluated result.

Responsibility and timing

Children finish independently. The Suite must retain NotEvaluated while Running, even when
a child is Failed, and wait for both child completion and helper completion before Completing.
The helper records the old child views; ProcessTestCases applies the next views afterwards.
Status counters must already reflect those new views in the same Suite call.

Isolation

Only the Suite subject publishes to the local capture. Child and helper doubles supply
controlled observations, not scheduling or lifecycle implementations. The test acts as parent
for the subject's own reservations and releases them at successful Reset and completion.
Detailed finalization and reservation-delegation checks belong to their dedicated scenarios.
</description>
*)
{endregion}
FUNCTION_BLOCK Test_SuiteNormalLifecycle EXTENDS TestCaseBase
VAR_INPUT
    FirstChildResult : E_Result := E_Result.Passed; //! Scenario parameter: Passed or Failed, held constant by the containing test Suite.
END_VAR
VAR
    FSubjectParent : I_RunControl;
    FSubject : TestSuiteLifecycleProbe;
    FHelper : SuiteOrchestratorDouble;
    FCapture : EventBuffer;
    FEvents : ARRAY[1..CaptureLength] OF ST_Event;
    FCaptureFifo : ST_FifoStatus;
    FCaptureStatus : ST_EventBufferStatus;
    FStep : INT;
    FStepChecked : BOOL;
    FStatePath : AssertTrue;
    FStatePathMatches : BOOL := TRUE;
    FTaskMapping : AssertTrue;
    FTaskMappingMatches : BOOL := TRUE;
    FOwnerResult : AssertTrue;
    FOwnerResultMatches : BOOL := TRUE;
    FStatusCounters : AssertTrue;
    FStatusCountersMatches : BOOL := TRUE;
    FCallOrder : AssertTrue;
    FCallOrderMatches : BOOL := TRUE;
    FReadiness : AssertTrue;
    FReadinessMatches : BOOL := TRUE;
    FCaptureIntegrity : AssertTrue;
    FCaptureIntegrityMatches : BOOL := TRUE;
END_VAR
VAR CONSTANT
    CaptureLength : UINT := 64;
    ChildCount : UINT := 2;
    Setup : INT := 0;
    ResetRequested : INT := 1;
    ChildrenReady : INT := 2;
    ResetFinished : INT := 3;
    StartReady : INT := 4;
    StartRequested : INT := 5;
    FirstChildCompleted : INT := 6;
    AllChildrenCompleted : INT := 7;
    WaitForHelper : INT := 8;
    OwnerCompleting : INT := 9;
    OwnerCompleted : INT := 10;
    StepCount : INT := 11;
END_VAR

SUPER^();

{region 'Documentation'}
(*!
<summary>Contributes only the checking Assertions, not the intentionally controlled subject results.</summary>
*)
{endregion}
METHOD PROTECTED AggregateResults
VAR_INPUT
    Aggregator : I_ResultAggregator; //! Borrowed result sink owned by the outer Test Case; add this test's checking Assertions without resetting or retaining the sink.
END_VAR
Aggregator.AddProvider(Provider := FStatePath);
Aggregator.AddProvider(Provider := FTaskMapping);
Aggregator.AddProvider(Provider := FOwnerResult);
Aggregator.AddProvider(Provider := FStatusCounters);
Aggregator.AddProvider(Provider := FCallOrder);
Aggregator.AddProvider(Provider := FReadiness);
Aggregator.AddProvider(Provider := FCaptureIntegrity);
END_METHOD

{region 'Documentation'}
(*!
<summary>Supplies only the root identity; the root never executes this isolated subject.</summary>
*)
{endregion}
METHOD PUBLIC BindSubjectParent
VAR_INPUT
    Parent : I_RunControl; //! Borrowed identity parent retained for isolated subject initialization; keep the Run-Control alive through subject use.
END_VAR
FSubjectParent := Parent;
END_METHOD

{region 'Documentation'}
(*!
<summary>Initializes the checking Assertions; the scenario explicitly initializes its isolated subject.</summary>
*)
{endregion}
METHOD PROTECTED Configure
FPreparationStateCount := 0;
FTestStateCount := StepCount;
FStatePath.Initialize(Parent := THIS^,
    AssertionName := 'StatePath');
FTaskMapping.Initialize(Parent := THIS^,
    AssertionName := 'TaskMapping');
FOwnerResult.Initialize(Parent := THIS^,
    AssertionName := 'OwnerResult');
FStatusCounters.Initialize(Parent := THIS^,
    AssertionName := 'StatusCounters');
FCallOrder.Initialize(Parent := THIS^,
    AssertionName := 'CallOrder');
FReadiness.Initialize(Parent := THIS^,
    AssertionName := 'Readiness');
FCaptureIntegrity.Initialize(Parent := THIS^,
    AssertionName := 'CaptureIntegrity');
END_METHOD

{region 'Documentation'}
(*!
<summary>No asynchronous test resource remains to stop.</summary>
*)
{endregion}
METHOD PROTECTED ProcessAbort
VAR_INPUT
    Enable : BOOL; //! Phase permission supplied by the owning Test Case; FALSE does not authorize progression, while observation may continue.
END_VAR
IF Enable THEN
    CompleteAbort();
END_IF;
END_METHOD

{region 'Documentation'}
(*!
<summary>Evaluates each step before advancing; assertions retain failures across the full owner lifecycle.</summary>
*)
{endregion}
METHOD PROTECTED ProcessAssertions
VAR_INPUT
    Enable : BOOL; //! Phase permission supplied by the owning Test Case; FALSE does not authorize progression, while observation may continue.
END_VAR
FStatePath(Enable := Enable,
    State := State,
    IN := FStatePathMatches);
FTaskMapping(Enable := Enable,
    State := State,
    IN := FTaskMappingMatches);
FOwnerResult(Enable := Enable,
    State := State,
    IN := FOwnerResultMatches);
FStatusCounters(Enable := Enable,
    State := State,
    IN := FStatusCountersMatches);
FCallOrder(Enable := Enable,
    State := State,
    IN := FCallOrderMatches);
FReadiness(Enable := Enable,
    State := State,
    IN := FReadinessMatches);
FCaptureIntegrity(Enable := Enable,
    State := State,
    IN := FCaptureIntegrityMatches);
IF Enable THEN
    FStepChecked := TRUE;
END_IF;
END_METHOD

{region 'Documentation'}
(*!
<summary>No resource Preparation is required for this controlled owner scenario.</summary>
*)
{endregion}
METHOD PROTECTED ProcessPreparations
VAR_INPUT
    // SA0033: Required override; the scenario has no Preparation phase.
    {attribute 'analysis' := '-33'}
    Enable : BOOL; //! Phase permission supplied by the owning Test Case; FALSE does not authorize progression, while observation may continue.
END_VAR
END_METHOD

{region 'Documentation'}
(*!
<summary>Restarts the test script and clears checking Assertions; subject setup belongs to the next test attempt.</summary>
*)
{endregion}
METHOD PROTECTED ProcessReset
FStep := Setup;
FStepChecked := FALSE;
FStatePathMatches := TRUE;
FTaskMappingMatches := TRUE;
FOwnerResultMatches := TRUE;
FStatusCountersMatches := TRUE;
FCallOrderMatches := TRUE;
FReadinessMatches := TRUE;
FCaptureIntegrityMatches := TRUE;
FStatePath.Reset();
FTaskMapping.Reset();
FOwnerResult.Reset();
FStatusCounters.Reset();
FCallOrder.Reset();
FReadiness.Reset();
FCaptureIntegrity.Reset();
CompleteReset();
END_METHOD

{region 'Documentation'}
(*!
<summary>Advances the explicit test script with at most one subject FB call per active PLC cycle.</summary>
*)
{endregion}
METHOD PROTECTED ProcessTests
VAR_INPUT
    Enable : BOOL; //! Phase permission supplied by the owning Test Case; FALSE does not authorize progression, while observation may continue.
END_VAR
IF NOT Enable THEN
    RETURN;
END_IF;
IF FStepChecked THEN
    IF FStep = OwnerCompleted THEN
        CompleteTests();
        RETURN;
    END_IF;
    FStep := FStep + 1;
    FStepChecked := FALSE;
    NextTestState();
END_IF;
RunStep();
END_METHOD

{region 'Documentation'}
(*!
<summary>Arranges one normal lifecycle cycle, executes the real Suite once, then records independent expectations.</summary>
*)
{endregion}
METHOD PRIVATE RunStep
VAR
    Config : ST_TestSuiteConfig;
    FirstView : ST_OrchestrationObservation;
    SecondView : ST_OrchestrationObservation;
    ExpectedState : E_State;
    ExpectedTask : E_OrchestratorTask;
    ExpectedResult : E_Result := E_Result.NotEvaluated;
    ExpectedReady : BOOL;
    ExpectedIdleCount : UINT;
    ExpectedRunningCount : UINT;
    ExpectedCompletedCount : UINT;
    ExpectedPassedCount : UINT;
    ExpectedFailedCount : UINT;
    ExpectedExecutionStatus : E_ExecutionStatus;
    FirstChild : I_Orchestratable;
    LastChild : I_Orchestratable;
    FirstStateBeforeCall : E_State;
    LastStateBeforeCall : E_State;
    Snapshot : ST_TestSuiteStatus;
END_VAR
CASE FStep OF
    Setup:
        IF NOT FCapture.Initialize(Buffer := FEvents,
            FifoControl := FCaptureFifo,
            Status := FCaptureStatus) THEN
            Error(Message := 'Suite lifecycle capture could not be initialized.');
            RETURN;
        END_IF;
        FHelper.BeginScenario();
        FSubject.Bind(Publisher := FCapture,
            Helper := FHelper);
        IF NOT FSubject.Initialize(Parent := FSubjectParent,
            SuiteName := 'LifecycleSubject',
            Config := Config) THEN
            Error(Message := 'Suite lifecycle subject could not be initialized.');
            RETURN;
        END_IF;
        FirstView.State := E_State.Uninitialized;
        FirstView.Ready := FALSE;
        SecondView := FirstView;
        ExpectedState := E_State.Uninitialized;
        ExpectedTask := E_OrchestratorTask.Idle;
        ExpectedExecutionStatus := E_ExecutionStatus.NotReady;

    ResetRequested:
        IF FSubject.ReserveResetEvents() <> E_EventReservationResult.Accepted THEN
            Error(Message := 'Suite lifecycle Reset reservation was rejected.');
            RETURN;
        END_IF;
        FSubject.RequestReset();
        FirstView.State := E_State.Reset;
        FirstView.Ready := FALSE;
        SecondView := FirstView;
        ExpectedState := E_State.Reset;
        ExpectedTask := E_OrchestratorTask.Reset;
        ExpectedExecutionStatus := E_ExecutionStatus.Reset;

    ChildrenReady:
        FSubject.RequestReset();
        ExpectedState := E_State.Reset;
        ExpectedTask := E_OrchestratorTask.Reset;
        ExpectedExecutionStatus := E_ExecutionStatus.Reset;
        ExpectedIdleCount := ChildCount;

    ResetFinished:
        FSubject.RequestReset();
        FHelper.SetObservation(Ready := FALSE,
            ResetFinished := TRUE);
        ExpectedState := E_State.Idle;
        ExpectedTask := E_OrchestratorTask.Idle;
        ExpectedExecutionStatus := E_ExecutionStatus.Idle;
        ExpectedIdleCount := ChildCount;

    StartReady:
        FHelper.SetObservation(Ready := TRUE);
        ExpectedState := E_State.Idle;
        ExpectedTask := E_OrchestratorTask.Idle;
        ExpectedExecutionStatus := E_ExecutionStatus.Idle;
        ExpectedIdleCount := ChildCount;
        ExpectedReady := TRUE;

    StartRequested:
        IF FSubject.ReserveExecutionEvents() <> E_EventReservationResult.Accepted THEN
            Error(Message := 'Suite lifecycle execution reservation was rejected.');
            RETURN;
        END_IF;
        FSubject.RequestStart();
        FirstView.State := E_State.Running;
        FirstView.Ready := FALSE;
        ExpectedState := E_State.Starting;
        ExpectedTask := E_OrchestratorTask.Execution;
        ExpectedExecutionStatus := E_ExecutionStatus.Starting;
        ExpectedIdleCount := 1;
        ExpectedRunningCount := 1;

    FirstChildCompleted:
        FHelper.SetObservation(Ready := FALSE);
        FirstView.State := E_State.Completed;
        FirstView.Result := FirstChildResult;
        FirstView.Ready := FALSE;
        FirstView.Complete := TRUE;
        SecondView.State := E_State.Running;
        SecondView.Ready := FALSE;
        ExpectedState := E_State.Running;
        ExpectedTask := E_OrchestratorTask.Execution;
        ExpectedExecutionStatus := E_ExecutionStatus.Running;
        ExpectedRunningCount := 1;
        ExpectedCompletedCount := 1;
        ExpectedFailedCount := BOOL_TO_UINT(FirstChildResult = E_Result.Failed);
        ExpectedPassedCount := 1 - ExpectedFailedCount;

    AllChildrenCompleted, WaitForHelper, OwnerCompleting, OwnerCompleted:
        FirstView.State := E_State.Completed;
        FirstView.Result := FirstChildResult;
        FirstView.Ready := FALSE;
        FirstView.Complete := TRUE;
        SecondView := FirstView;
        SecondView.Result := E_Result.Passed;
        ExpectedTask := E_OrchestratorTask.Execution;
        ExpectedCompletedCount := ChildCount;
        ExpectedFailedCount := BOOL_TO_UINT(FirstChildResult = E_Result.Failed);
        ExpectedPassedCount := ChildCount - ExpectedFailedCount;
        CASE FStep OF
            AllChildrenCompleted, WaitForHelper:
                ExpectedState := E_State.Running;
                ExpectedExecutionStatus := E_ExecutionStatus.Running;
            OwnerCompleting:
                FHelper.SetObservation(Ready := FALSE,
                    ExecutionFinished := TRUE);
                ExpectedState := E_State.Completing;
                ExpectedExecutionStatus := E_ExecutionStatus.Completing;
                ExpectedResult := FirstChildResult;
            OwnerCompleted:
                ExpectedState := E_State.Completed;
                ExpectedTask := E_OrchestratorTask.Idle;
                ExpectedExecutionStatus := E_ExecutionStatus.Completed;
                ExpectedResult := FirstChildResult;
        ELSE
            Error(Message := 'Unexpected normal completion step.');
            RETURN;
        END_CASE;
ELSE
    Error(Message := 'Unexpected Suite lifecycle test step.');
    RETURN;
END_CASE;

FirstChild := FSubject.GetChild(Index := FSubject.ChildArrayLowerBound);
LastChild := FSubject.GetChild(Index := FSubject.ChildArrayLowerBound + UINT_TO_DINT(FSubject.ChildCount) - 1);
FirstStateBeforeCall := FirstChild.State;
LastStateBeforeCall := LastChild.State;
FSubject.SetChildObservations(FirstChild := FirstView,
    SecondChild := SecondView);
FSubject();
Snapshot := FSubject.Status;

FStatePathMatches := (FSubject.State = ExpectedState)
    AND (Snapshot.Execution.State = ExpectedState)
    AND (Snapshot.Execution.ExecutionStatus = ExpectedExecutionStatus);
FTaskMappingMatches := FHelper.CurrentTask = ExpectedTask;
FOwnerResultMatches := (FSubject.Result = ExpectedResult)
    AND (Snapshot.Execution.Result = ExpectedResult)
    AND NOT FSubject.HasError;
FStatusCountersMatches := (Snapshot.TestCaseCountTotal = ChildCount)
    AND (Snapshot.TestCaseCountIdle = ExpectedIdleCount)
    AND (Snapshot.TestCaseCountRunning = ExpectedRunningCount)
    AND (Snapshot.TestCaseCountCompleted = ExpectedCompletedCount)
    AND (Snapshot.TestCaseCountPassed = ExpectedPassedCount)
    AND (Snapshot.TestCaseCountFailed = ExpectedFailedCount)
    AND (Snapshot.TestCaseCountError = 0) AND (Snapshot.TestCaseCountInactive = 0);
FCallOrderMatches := (FHelper.InitializeCount = 1)
    AND (FHelper.ExecuteCount = INT_TO_UINT(FStep + 1))
    AND (FSubject.ChildCallCount = INT_TO_UINT(FStep + 1))
    AND FSubject.ChildBodyCallsMatch
    AND (FHelper.FirstChildStateAtExecute = FirstStateBeforeCall)
    AND (FHelper.LastChildStateAtExecute = LastStateBeforeCall)
    AND (FirstChild.State = FirstView.State) AND (LastChild.State = SecondView.State);
FReadinessMatches := (FSubject.IsReady = ExpectedReady)
    AND (Snapshot.Execution.Ready = ExpectedReady)
    AND (FSubject.IsComplete = (ExpectedState = E_State.Completed));
FCaptureIntegrityMatches := FCaptureStatus.LostEventCount = 0;

IF (FStep = ResetFinished) OR (FStep = OwnerCompleted) THEN
    IF NOT FSubject.FreeReservedEvents() THEN
        Error(Message := 'Suite lifecycle fixture could not release its reservation.');
    END_IF;
END_IF;
END_METHOD

END_FUNCTION_BLOCK

// ---- SelfTests/TestCases/TestSuite_TestSuiteLifecycle/Test_SuiteExceptionalLifecycle.TcPOU
{region 'Documentation'}
(*!
<summary>Exercises Suite error and Abort paths through controlled child/helper observations.</summary>
<description>

Scenario ownership

Each instance runs one selected scenario. Production Suite sequencing, timers, result handling
and publication stay unchanged. The local helper supplies observations, never child scheduling.
Only the isolated subject writes to the local capture; checking Assertions use the normal publisher.

Script and call order

RunStep arranges one cycle, calls the subject once, then checks the expected owner response.
FNextStep is accepted only after checking Assertions ran. Child snapshots are applied by the
subject's ProcessTestCases, so child errors affect the result in that call and the next Sequencer call.

Timeout and recovery

The three timeout scenarios withhold completion for the real configured deadline. Waiting
repeats a checkpoint, not subject calls within a cycle. The outer Test Case timeout bounds a
missing transition. These tests check the reaction and retained flags, not exact clock precision.
ResetTimeout submits another Reset on every waiting call, including the expired-deadline call.
The error scenario repeats Reset while Error is held and when the helper finally completes.
Every scenario ends with a successful lifecycle Reset without replacing bindings or configuration;
a scripted previous helper Error must not leak through the first-entry sequencing boundary.
</description>
*)
{endregion}
FUNCTION_BLOCK Test_SuiteExceptionalLifecycle EXTENDS TestCaseBase
VAR_INPUT
    Scenario : E_SuiteLifecycleScenario := E_SuiteLifecycleScenario.ResetError; //! Fixed scenario selection supplied by the containing Suite on every call.
END_VAR
VAR
    FSubjectParent : I_RunControl;
    FSubject : TestSuiteLifecycleProbe;
    FHelper : SuiteOrchestratorDouble;
    FCapture : EventBuffer;
    FEvents : ARRAY[1..CaptureLength] OF ST_Event;
    FCaptureFifo : ST_FifoStatus;
    FCaptureStatus : ST_EventBufferStatus;
    FFirstChild : ST_OrchestrationObservation;
    FSecondChild : ST_OrchestrationObservation;
    FStep : INT;
    FNextStep : INT;
    FStepChecked : BOOL;
    FSubjectCallCount : UINT;
    FExpectedTimeout : BOOL;
    FExpectedResetTimeout : BOOL;
    FExpectedAbortTimeout : BOOL;
    FStatePath : AssertTrue;
    FStatePathMatches : BOOL := TRUE;
    FTaskMapping : AssertTrue;
    FTaskMappingMatches : BOOL := TRUE;
    FResultStatus : AssertTrue;
    FResultStatusMatches : BOOL := TRUE;
    FTimeoutFlags : AssertTrue;
    FTimeoutFlagsMatches : BOOL := TRUE;
    FChildCalls : AssertTrue;
    FChildCallsMatches : BOOL := TRUE;
    FDiagnostics : AssertTrue;
    FDiagnosticsMatches : BOOL := TRUE;
    FRecovery : AssertTrue;
    FRecoveryMatches : BOOL := TRUE;
END_VAR
VAR CONSTANT
    CaptureLength : UINT := 128;
    ShortTimeout : TIME := T#50ms;
    Setup : INT := 0;
    RequestInitialReset : INT := 1;
    InitialResetResponse : INT := 2;
    HoldResetError : INT := 3;
    FinishFailedReset : INT := 4;
    StartExecution : INT := 5;
    ReachRunning : INT := 6;
    ApplyStimulus : INT := 7;
    ObserveChildError : INT := 8;
    ObserveAbortResponse : INT := 9;
    FinishChildren : INT := 10;
    FinishHelper : INT := 11;
    CheckCompleted : INT := 12;
    RecoveryReset : INT := 13;
    RecoveryReady : INT := 14;
    Done : INT := 15;
END_VAR

SUPER^();

{region 'Documentation'}
(*!
<summary>Contributes only the checking Assertions, not the intentionally controlled subject results.</summary>
*)
{endregion}
METHOD PROTECTED AggregateResults
VAR_INPUT
    Aggregator : I_ResultAggregator; //! Borrowed result sink owned by the outer Test Case; add this test's checking Assertions without resetting or retaining the sink.
END_VAR
Aggregator.AddProvider(Provider := FStatePath);
Aggregator.AddProvider(Provider := FTaskMapping);
Aggregator.AddProvider(Provider := FResultStatus);
Aggregator.AddProvider(Provider := FTimeoutFlags);
Aggregator.AddProvider(Provider := FChildCalls);
Aggregator.AddProvider(Provider := FDiagnostics);
Aggregator.AddProvider(Provider := FRecovery);
END_METHOD

{region 'Documentation'}
(*!
<summary>Supplies only the root identity; the root never executes this isolated subject.</summary>
*)
{endregion}
METHOD PUBLIC BindSubjectParent
VAR_INPUT
    Parent : I_RunControl; //! Borrowed identity parent retained for isolated subject initialization; keep the Run-Control alive through subject use.
END_VAR
FSubjectParent := Parent;
END_METHOD

{region 'Documentation'}
(*!
<summary>Checks structured owner diagnostics and forbids Abort transitions for failed Reset; ignores message wording.</summary>
*)
{endregion}
METHOD PRIVATE CheckDiagnostics
VAR
    Index : UINT;
    DiagnosticCount : UINT;
    AbortTransitionCount : UINT;
END_VAR
FOR Index := 1 TO CaptureLength DO
    IF (FEvents[Index].SequenceId = 0) OR (FEvents[Index].Name <> FSubject.Name) THEN
        CONTINUE;
    END_IF;
    IF (FEvents[Index].EventType = E_EventType.Framework)
        AND (FEvents[Index].Severity = E_EventSeverity.Error) THEN
        DiagnosticCount := DiagnosticCount + 1;
    END_IF;
    IF (FEvents[Index].EventType = E_EventType.StateTransition)
        AND ((FEvents[Index].State = E_State.Aborting)
            OR (FEvents[Index].State = E_State.AbortingFromError)) THEN
        AbortTransitionCount := AbortTransitionCount + 1;
    END_IF;
END_FOR;
IF Scenario = E_SuiteLifecycleScenario.Abort THEN
    FDiagnosticsMatches := DiagnosticCount = 0;
ELSE
    FDiagnosticsMatches := DiagnosticCount = 1;
END_IF;
IF (Scenario = E_SuiteLifecycleScenario.ResetError) OR (Scenario = E_SuiteLifecycleScenario.ResetTimeout) THEN
    FDiagnosticsMatches := FDiagnosticsMatches AND (AbortTransitionCount = 0);
ELSE
    FDiagnosticsMatches := FDiagnosticsMatches AND (AbortTransitionCount > 0);
END_IF;
FDiagnosticsMatches := FDiagnosticsMatches AND (FCaptureStatus.LostEventCount = 0);
END_METHOD

{region 'Documentation'}
(*!
<summary>Initializes the checking Assertions; the scenario explicitly initializes its isolated subject.</summary>
*)
{endregion}
METHOD PROTECTED Configure
FPreparationStateCount := 0;
FTestStateCount := 1;
FStatePath.Initialize(Parent := THIS^,
    AssertionName := 'StatePath');
FTaskMapping.Initialize(Parent := THIS^,
    AssertionName := 'TaskMapping');
FResultStatus.Initialize(Parent := THIS^,
    AssertionName := 'ResultStatus');
FTimeoutFlags.Initialize(Parent := THIS^,
    AssertionName := 'TimeoutFlags');
FChildCalls.Initialize(Parent := THIS^,
    AssertionName := 'ChildCalls');
FDiagnostics.Initialize(Parent := THIS^,
    AssertionName := 'Diagnostics');
FRecovery.Initialize(Parent := THIS^,
    AssertionName := 'Recovery');
END_METHOD

{region 'Documentation'}
(*!
<summary>No asynchronous test resource remains to stop.</summary>
*)
{endregion}
METHOD PROTECTED ProcessAbort
VAR_INPUT
    Enable : BOOL; //! Phase permission supplied by the owning Test Case; FALSE does not authorize progression, while observation may continue.
END_VAR
IF Enable THEN
    CompleteAbort();
END_IF;
END_METHOD

{region 'Documentation'}
(*!
<summary>Checks every subject cycle before advancing, retaining failures across waiting and recovery.</summary>
*)
{endregion}
METHOD PROTECTED ProcessAssertions
VAR_INPUT
    Enable : BOOL; //! Phase permission supplied by the owning Test Case; FALSE does not authorize progression, while observation may continue.
END_VAR
FStatePath(Enable := Enable,
    State := State,
    IN := FStatePathMatches);
FTaskMapping(Enable := Enable,
    State := State,
    IN := FTaskMappingMatches);
FResultStatus(Enable := Enable,
    State := State,
    IN := FResultStatusMatches);
FTimeoutFlags(Enable := Enable,
    State := State,
    IN := FTimeoutFlagsMatches);
FChildCalls(Enable := Enable,
    State := State,
    IN := FChildCallsMatches);
FDiagnostics(Enable := Enable,
    State := State,
    IN := FDiagnosticsMatches);
FRecovery(Enable := Enable,
    State := State,
    IN := FRecoveryMatches);
IF Enable THEN
    FStepChecked := TRUE;
END_IF;
END_METHOD

{region 'Documentation'}
(*!
<summary>No resource Preparation is required for this controlled owner scenario.</summary>
*)
{endregion}
METHOD PROTECTED ProcessPreparations
VAR_INPUT
    // SA0033: Required override; the scenario has no Preparation phase.
    {attribute 'analysis' := '-33'}
    Enable : BOOL; //! Phase permission supplied by the owning Test Case; FALSE does not authorize progression, while observation may continue.
END_VAR
END_METHOD

{region 'Documentation'}
(*!
<summary>Restarts the test script and clears checking Assertions; subject setup belongs to the next test attempt.</summary>
*)
{endregion}
METHOD PROTECTED ProcessReset
FStep := Setup;
FNextStep := Setup;
FStepChecked := FALSE;
FSubjectCallCount := 0;
FExpectedTimeout := FALSE;
FExpectedResetTimeout := FALSE;
FExpectedAbortTimeout := FALSE;
FStatePathMatches := TRUE;
FTaskMappingMatches := TRUE;
FResultStatusMatches := TRUE;
FTimeoutFlagsMatches := TRUE;
FChildCallsMatches := TRUE;
FDiagnosticsMatches := TRUE;
FRecoveryMatches := TRUE;
FStatePath.Reset();
FTaskMapping.Reset();
FResultStatus.Reset();
FTimeoutFlags.Reset();
FChildCalls.Reset();
FDiagnostics.Reset();
FRecovery.Reset();
CompleteReset();
END_METHOD

{region 'Documentation'}
(*!
<summary>Advances the explicit test script with at most one subject FB call per active PLC cycle.</summary>
*)
{endregion}
METHOD PROTECTED ProcessTests
VAR_INPUT
    Enable : BOOL; //! Phase permission supplied by the owning Test Case; FALSE does not authorize progression, while observation may continue.
END_VAR
IF NOT Enable THEN
    RETURN;
END_IF;
IF FStepChecked THEN
    FStep := FNextStep;
    FStepChecked := FALSE;
END_IF;
IF FStep = Done THEN
    CompleteTests();
    RETURN;
END_IF;
RunStep();
END_METHOD

{region 'Documentation'}
(*!
<summary>Arranges one error-path checkpoint and checks the real Suite; timeout waits use further PLC cycles.</summary>
*)
{endregion}
METHOD PRIVATE RunStep
VAR
    Config : ST_TestSuiteConfig;
    Snapshot : ST_TestSuiteStatus;
    ExpectedState : E_State;
    ExpectedTask : E_OrchestratorTask;
    ExpectedResult : E_Result;
    FinalResult : E_Result;
    WaitForTimeout : BOOL;
    WaitingState : E_State;
    WaitingTask : E_OrchestratorTask;
    WaitingResult : E_Result := E_Result.NotEvaluated;
END_VAR
FNextStep := FStep + 1;
ExpectedResult := E_Result.NotEvaluated;
ExpectedTask := E_OrchestratorTask.Idle;
FinalResult := E_Result.Error;
IF Scenario = E_SuiteLifecycleScenario.Abort THEN
    FinalResult := E_Result.Abort;
END_IF;

CASE FStep OF
    Setup:
        CASE Scenario OF
            E_SuiteLifecycleScenario.ResetTimeout:
                Config.ResetTimeout := ShortTimeout;
            E_SuiteLifecycleScenario.ExecutionTimeout:
                Config.Timeout := ShortTimeout;
            E_SuiteLifecycleScenario.AbortTimeout:
                Config.AbortTimeout := ShortTimeout;
        ELSE
            // Other scenarios use the ordinary positive deadlines.
        END_CASE;
        IF NOT FCapture.Initialize(Buffer := FEvents,
            FifoControl := FCaptureFifo,
            Status := FCaptureStatus) THEN
            Error(Message := 'Exceptional Suite capture could not be initialized.');
            RETURN;
        END_IF;
        FHelper.BeginScenario();
        FSubject.Bind(Publisher := FCapture,
            Helper := FHelper);
        IF NOT FSubject.Initialize(Parent := FSubjectParent,
            SuiteName := 'ExceptionalSubject',
            Config := Config) THEN
            Error(Message := 'Exceptional Suite subject could not be initialized.');
            RETURN;
        END_IF;
        FFirstChild.State := E_State.Uninitialized;
        FFirstChild.Result := E_Result.NotEvaluated;
        FFirstChild.Ready := FALSE;
        FFirstChild.Complete := FALSE;
        FSecondChild := FFirstChild;
        ExpectedState := E_State.Uninitialized;

    RequestInitialReset:
        IF FSubject.ReserveResetEvents() <> E_EventReservationResult.Accepted THEN
            Error(Message := 'Initial Suite Reset reservation was rejected.');
            RETURN;
        END_IF;
        FSubject.RequestReset();
        FFirstChild.State := E_State.Reset;
        FSecondChild := FFirstChild;
        ExpectedState := E_State.Reset;
        ExpectedTask := E_OrchestratorTask.Reset;

    InitialResetResponse:
        CASE Scenario OF
            E_SuiteLifecycleScenario.ResetError:
                FHelper.SetObservation(Ready := FALSE,
                    Result := E_Result.Error);
                FFirstChild.State := E_State.Completed;
                FFirstChild.Result := E_Result.Error;
                FFirstChild.Complete := TRUE;
                ExpectedState := E_State.Reset;
                ExpectedResult := E_Result.Error;
                ExpectedTask := E_OrchestratorTask.Reset;
                FNextStep := HoldResetError;

            E_SuiteLifecycleScenario.ResetTimeout:
                FSubject.RequestReset();
                WaitForTimeout := TRUE;
                WaitingState := E_State.Reset;
                WaitingTask := E_OrchestratorTask.Reset;
                ExpectedState := E_State.Completing;
                ExpectedResult := E_Result.Error;
                FNextStep := CheckCompleted;
        ELSE
            FHelper.SetObservation(Ready := TRUE,
                ResetFinished := TRUE);
            FFirstChild.State := E_State.Idle;
            FFirstChild.Ready := TRUE;
            FSecondChild := FFirstChild;
            ExpectedState := E_State.Idle;
            FNextStep := StartExecution;
        END_CASE;

    HoldResetError:
        // Another Reset request must not clear the held error or abandon the unfinished child.
        FSubject.RequestReset();
        ExpectedState := E_State.Reset;
        ExpectedResult := E_Result.Error;
        ExpectedTask := E_OrchestratorTask.Reset;

    FinishFailedReset:
        FSubject.RequestReset();
        FHelper.SetObservation(Ready := FALSE,
            Result := E_Result.Error,
            ResetFinished := TRUE);
        FSecondChild.State := E_State.Idle;
        FSecondChild.Ready := TRUE;
        ExpectedState := E_State.Completing;
        ExpectedResult := E_Result.Error;
        FNextStep := CheckCompleted;

    StartExecution:
        IF FSubject.ReserveExecutionEvents() <> E_EventReservationResult.Accepted THEN
            Error(Message := 'Exceptional Suite execution reservation was rejected.');
            RETURN;
        END_IF;
        FSubject.RequestStart();
        FFirstChild.State := E_State.Running;
        FFirstChild.Ready := FALSE;
        ExpectedState := E_State.Starting;
        ExpectedTask := E_OrchestratorTask.Execution;

    ReachRunning:
        FHelper.SetObservation(Ready := FALSE);
        ExpectedState := E_State.Running;
        ExpectedTask := E_OrchestratorTask.Execution;

    ApplyStimulus:
        CASE Scenario OF
            E_SuiteLifecycleScenario.ChildError, E_SuiteLifecycleScenario.UnexpectedChildAbort:
                FFirstChild.State := E_State.Completed;
                FFirstChild.Complete := TRUE;
                IF Scenario = E_SuiteLifecycleScenario.ChildError THEN
                    FFirstChild.Result := E_Result.Error;
                ELSE
                    FFirstChild.Result := E_Result.Abort;
                END_IF;
                ExpectedState := E_State.Running;
                ExpectedResult := E_Result.Error;
                ExpectedTask := E_OrchestratorTask.Execution;
                FNextStep := ObserveChildError;

            E_SuiteLifecycleScenario.ExecutionError:
                FHelper.SetObservation(Ready := FALSE,
                    Result := E_Result.Error);
                ExpectedState := E_State.AbortingFromError;
                ExpectedResult := E_Result.Error;
                ExpectedTask := E_OrchestratorTask.Abort;
                FNextStep := FinishChildren;

            E_SuiteLifecycleScenario.ExecutionTimeout:
                WaitForTimeout := TRUE;
                WaitingState := E_State.Running;
                WaitingTask := E_OrchestratorTask.Execution;
                ExpectedState := E_State.AbortingFromError;
                ExpectedResult := E_Result.Error;
                ExpectedTask := E_OrchestratorTask.Abort;
                FNextStep := FinishChildren;

            E_SuiteLifecycleScenario.Abort, E_SuiteLifecycleScenario.AbortError, E_SuiteLifecycleScenario.AbortTimeout:
                FSubject.RequestAbort();
                FFirstChild.State := E_State.Aborting;
                FFirstChild.Result := E_Result.Abort;
                ExpectedState := E_State.Aborting;
                ExpectedResult := E_Result.Abort;
                ExpectedTask := E_OrchestratorTask.Abort;
                FNextStep := ObserveAbortResponse;
        ELSE
            Error(Message := 'Unsupported execution stimulus.');
            RETURN;
        END_CASE;

    ObserveChildError:
        ExpectedState := E_State.AbortingFromError;
        ExpectedResult := E_Result.Error;
        ExpectedTask := E_OrchestratorTask.Abort;
        FNextStep := FinishChildren;

    ObserveAbortResponse:
        CASE Scenario OF
            E_SuiteLifecycleScenario.Abort:
                ExpectedState := E_State.Aborting;
                ExpectedResult := E_Result.Abort;
                ExpectedTask := E_OrchestratorTask.Abort;
                FNextStep := FinishChildren;
            E_SuiteLifecycleScenario.AbortError:
                FHelper.SetObservation(Ready := FALSE,
                    Result := E_Result.Error);
                ExpectedState := E_State.AbortingFromError;
                ExpectedResult := E_Result.Error;
                ExpectedTask := E_OrchestratorTask.Abort;
                FNextStep := FinishChildren;
            E_SuiteLifecycleScenario.AbortTimeout:
                WaitForTimeout := TRUE;
                WaitingState := E_State.Aborting;
                WaitingResult := E_Result.Abort;
                WaitingTask := E_OrchestratorTask.Abort;
                ExpectedState := E_State.Completing;
                ExpectedResult := E_Result.Error;
                ExpectedTask := E_OrchestratorTask.Abort;
                FNextStep := CheckCompleted;
        ELSE
            Error(Message := 'Unsupported Abort observation.');
            RETURN;
        END_CASE;

    FinishChildren:
        FFirstChild.State := E_State.Completed;
        FFirstChild.Ready := FALSE;
        FFirstChild.Complete := TRUE;
        IF Scenario <> E_SuiteLifecycleScenario.ChildError THEN
            FFirstChild.Result := E_Result.Abort;
        END_IF;
        ExpectedState := E_State.AbortingFromError;
        IF Scenario = E_SuiteLifecycleScenario.Abort THEN
            ExpectedState := E_State.Aborting;
        END_IF;
        ExpectedResult := FinalResult;
        ExpectedTask := E_OrchestratorTask.Abort;

    FinishHelper:
        FHelper.SetObservation(Ready := FALSE,
            Result := FHelper.Result,
            AbortFinished := TRUE);
        ExpectedState := E_State.Completing;
        ExpectedResult := FinalResult;
        ExpectedTask := E_OrchestratorTask.Abort;

    CheckCompleted:
        ExpectedState := E_State.Completed;
        ExpectedResult := FinalResult;

    RecoveryReset:
        // Keep the previous task Error observable until the new helper task has been assigned.
        FHelper.SetObservation(Ready := FALSE,
            Result := E_Result.Error);
        IF FSubject.ReserveResetEvents() <> E_EventReservationResult.Accepted THEN
            Error(Message := 'Recovery Reset reservation was rejected.');
            RETURN;
        END_IF;
        FSubject.RequestReset();
        FFirstChild.State := E_State.Reset;
        FFirstChild.Result := E_Result.NotEvaluated;
        FFirstChild.Complete := FALSE;
        FFirstChild.Ready := FALSE;
        FSecondChild := FFirstChild;
        FExpectedTimeout := FALSE;
        FExpectedResetTimeout := FALSE;
        FExpectedAbortTimeout := FALSE;
        ExpectedState := E_State.Reset;
        ExpectedTask := E_OrchestratorTask.Reset;

    RecoveryReady:
        FHelper.SetObservation(Ready := TRUE,
            ResetFinished := TRUE);
        FFirstChild.State := E_State.Idle;
        FFirstChild.Ready := TRUE;
        FSecondChild := FFirstChild;
        ExpectedState := E_State.Idle;
ELSE
    Error(Message := 'Unexpected exceptional Suite test step.');
    RETURN;
END_CASE;

FSubject.SetChildObservations(FirstChild := FFirstChild,
    SecondChild := FSecondChild);
FSubject();
FSubjectCallCount := FSubjectCallCount + 1;
Snapshot := FSubject.Status;

IF WaitForTimeout THEN
    IF FSubject.State = WaitingState THEN
        ExpectedState := WaitingState;
        ExpectedTask := WaitingTask;
        ExpectedResult := WaitingResult;
        FNextStep := FStep;
    ELSE
        CASE Scenario OF
            E_SuiteLifecycleScenario.ResetTimeout:
                FExpectedResetTimeout := TRUE;
            E_SuiteLifecycleScenario.ExecutionTimeout:
                FExpectedTimeout := TRUE;
            E_SuiteLifecycleScenario.AbortTimeout:
                FExpectedAbortTimeout := TRUE;
        ELSE
            Error(Message := 'Unexpected timeout-wait scenario.');
            RETURN;
        END_CASE;
    END_IF;
END_IF;

FStatePathMatches := (FSubject.State = ExpectedState) AND (Snapshot.Execution.State = ExpectedState);
FTaskMappingMatches := FHelper.CurrentTask = ExpectedTask;
FResultStatusMatches := (FSubject.Result = ExpectedResult)
    AND (Snapshot.Execution.Result = ExpectedResult)
    AND (FSubject.HasError = (ExpectedResult = E_Result.Error))
    AND (Snapshot.Execution.Error = (ExpectedResult = E_Result.Error))
    AND (FSubject.IsComplete = (ExpectedState = E_State.Completed))
    AND (Snapshot.Execution.Completed = (ExpectedState = E_State.Completed));
FTimeoutFlagsMatches := (FSubject.HasTimeout = FExpectedTimeout)
    AND (FSubject.HasResetTimeout = FExpectedResetTimeout)
    AND (FSubject.HasAbortTimeout = FExpectedAbortTimeout);
FChildCallsMatches := (FHelper.ExecuteCount = FSubjectCallCount)
    AND (FSubject.ChildCallCount = FSubjectCallCount)
    AND FSubject.ChildBodyCallsMatch;

IF FStep = CheckCompleted THEN
    CheckDiagnostics();
END_IF;
IF (FStep = CheckCompleted) OR (FStep = RecoveryReady)
    OR ((FStep = InitialResetResponse) AND (ExpectedState = E_State.Idle)) THEN
    IF NOT FSubject.FreeReservedEvents() THEN
        Error(Message := 'Exceptional Suite fixture could not release its reservation.');
    END_IF;
END_IF;
IF FStep = RecoveryReady THEN
    FRecoveryMatches := FSubject.IsReady AND Snapshot.Execution.Ready
        AND (FSubject.Result = E_Result.NotEvaluated)
        AND (FHelper.InitializeCount = 1) AND (FSubject.ConfigureCount = 1)
        AND (FSubject.ReservedEntryCount = 0) AND (FCapture.ReservedEntryCount = 0)
        AND (FCaptureStatus.LostEventCount = 0);
END_IF;
END_METHOD

END_FUNCTION_BLOCK

// ---- SelfTests/TestCases/TestSuite_TestSuiteLifecycle/Test_SuiteFinalization.TcPOU
{region 'Documentation'}
(*!
<summary>Checks Suite finalization and ongoing observation with normal completion or late children after Reset timeout.</summary>
<description>

Publication boundary

The local capture must contain one Result and one Aggregation in Completing, followed by
the Completed transition on a later subject call. Exact payloads are retained for comparison.
The expected aggregation text is constructed from fixed scenario counts and observed runtime,
not through the production event constructor.

Late child observation

In the Reset-timeout variant the Suite completes while its children are still resetting.
One then reaches Completed/Error and the other Idle. The Suite must refresh its counters
without rewriting final events or restarting orchestration. The normal variant keeps both
children completed and verifies quiet repeated calls and synchronous reservation cleanup.
</description>
*)
{endregion}
FUNCTION_BLOCK Test_SuiteFinalization EXTENDS TestCaseBase
VAR_INPUT
    LateResetChildren : BOOL := FALSE; //! FALSE: normal Passed completion; TRUE: Reset timeout followed by delayed child completion.
END_VAR
VAR
    FSubjectParent : I_RunControl;
    FSubject : TestSuiteLifecycleProbe;
    FHelper : SuiteOrchestratorDouble;
    FCapture : EventBuffer;
    FEvents : ARRAY[1..CaptureLength] OF ST_Event;
    FCaptureFifo : ST_FifoStatus;
    FCaptureStatus : ST_EventBufferStatus;
    FFirstChild : ST_OrchestrationObservation;
    FSecondChild : ST_OrchestrationObservation;
    FStep : INT;
    FNextStep : INT;
    FStepChecked : BOOL;
    FSubjectCalls : UINT;
    FExpectFinalization : BOOL;
    FExpectCompletion : BOOL;
    FSavedFinalization : BOOL;
    FFinalizationCall : UINT;
    FExpectedFinalResult : E_Result;
    FResultSnapshot : ST_Event;
    FAggregationSnapshot : ST_Event;
    FExpectedAggregation : STRING(GVL_Constants.MessageLength);
    FCompletedSequence : UDINT;
    FLifecycle : AssertTrue;
    FLifecycleMatches : BOOL := TRUE;
    FPublication : AssertTrue;
    FPublicationMatches : BOOL := TRUE;
    FEventOrder : AssertTrue;
    FEventOrderMatches : BOOL := TRUE;
    FFrozenPayload : AssertTrue;
    FFrozenPayloadMatches : BOOL := TRUE;
    FStatusRefresh : AssertTrue;
    FStatusRefreshMatches : BOOL := TRUE;
    FChildCalls : AssertTrue;
    FChildCallsMatches : BOOL := TRUE;
    FCleanup : AssertTrue;
    FCleanupMatches : BOOL := TRUE;
END_VAR
VAR CONSTANT
    CaptureLength : UINT := 64;
    Setup : INT := 0;
    ResetRequested : INT := 1;
    ResetOutcome : INT := 2;
    StartRequested : INT := 3;
    CompleteChildren : INT := 4;
    CompleteOwner : INT := 5;
    CompleteState : INT := 6;
    LateChildProgress : INT := 7;
    QuietCompleted : INT := 8;
    ReleaseReservations : INT := 9;
    QuietAfterRelease : INT := 10;
    Done : INT := 11;
END_VAR

SUPER^();

{region 'Documentation'}
(*!
<summary>Contributes only the checking Assertions, not the intentionally controlled subject results.</summary>
*)
{endregion}
METHOD PROTECTED AggregateResults
VAR_INPUT
    Aggregator : I_ResultAggregator; //! Borrowed result sink owned by the outer Test Case; add this test's checking Assertions without resetting or retaining the sink.
END_VAR
Aggregator.AddProvider(Provider := FLifecycle);
Aggregator.AddProvider(Provider := FPublication);
Aggregator.AddProvider(Provider := FEventOrder);
Aggregator.AddProvider(Provider := FFrozenPayload);
Aggregator.AddProvider(Provider := FStatusRefresh);
Aggregator.AddProvider(Provider := FChildCalls);
Aggregator.AddProvider(Provider := FCleanup);
END_METHOD

{region 'Documentation'}
(*!
<summary>Supplies only the root identity; the root never executes this isolated subject.</summary>
*)
{endregion}
METHOD PUBLIC BindSubjectParent
VAR_INPUT
    Parent : I_RunControl; //! Borrowed identity parent retained for isolated subject initialization; keep the Run-Control alive through subject use.
END_VAR
FSubjectParent := Parent;
END_METHOD

{region 'Documentation'}
(*!
<summary>Counts owner finalization events and checks original payloads and order without consuming the capture.</summary>
*)
{endregion}
METHOD PRIVATE CheckEventStream
VAR
    Index : UINT;
    ResultIndex : UINT;
    AggregationIndex : UINT;
    ResultCount : UINT;
    AggregationCount : UINT;
    CompletionCount : UINT;
    CompletionSequence : UDINT;
END_VAR
FOR Index := 1 TO CaptureLength DO
    IF (FEvents[Index].SequenceId = 0) OR (FEvents[Index].Name <> FSubject.Name) THEN
        CONTINUE;
    END_IF;
    CASE FEvents[Index].EventType OF
        E_EventType.Result:
            ResultCount := ResultCount + 1;
            ResultIndex := Index;
        E_EventType.Aggregation:
            AggregationCount := AggregationCount + 1;
            AggregationIndex := Index;
        E_EventType.StateTransition:
            IF FEvents[Index].State = E_State.Completed THEN
                CompletionCount := CompletionCount + 1;
                CompletionSequence := FEvents[Index].SequenceId;
            END_IF;
    ELSE
        // Triggers and diagnostics are not finalization events.
    END_CASE;
END_FOR;
FPublicationMatches := (ResultCount = BOOL_TO_UINT(FExpectFinalization))
    AND (AggregationCount = BOOL_TO_UINT(FExpectFinalization))
    AND (CompletionCount = BOOL_TO_UINT(FExpectCompletion))
    AND (FCaptureStatus.LostEventCount = 0);
IF NOT FExpectFinalization OR (ResultCount <> 1) OR (AggregationCount <> 1) THEN
    RETURN;
END_IF;

FPublicationMatches := FPublicationMatches
    AND (FEvents[ResultIndex].OwnerScope = E_OwnerScope.TestSuite)
    AND (FEvents[AggregationIndex].OwnerScope = E_OwnerScope.TestSuite)
    AND (FEvents[ResultIndex].State = E_State.Completing)
    AND (FEvents[AggregationIndex].State = E_State.Completing)
    AND (FEvents[ResultIndex].Result = FExpectedFinalResult)
    AND (FEvents[AggregationIndex].Result = FExpectedFinalResult)
    AND (FEvents[AggregationIndex].Message = FExpectedAggregation);
FEventOrderMatches := FEvents[ResultIndex].SequenceId < FEvents[AggregationIndex].SequenceId;
IF NOT FSavedFinalization THEN
    FResultSnapshot := FEvents[ResultIndex];
    FAggregationSnapshot := FEvents[AggregationIndex];
    FFinalizationCall := FSubjectCalls;
    FSavedFinalization := TRUE;
    FEventOrderMatches := FEventOrderMatches AND (FSubject.State = E_State.Completing);
END_IF;
IF FExpectCompletion THEN
    FEventOrderMatches := FEventOrderMatches
        AND (FEvents[AggregationIndex].SequenceId < CompletionSequence)
        AND (FSubjectCalls > FFinalizationCall);
END_IF;
FFrozenPayloadMatches := IsEventUnchanged(Event := FEvents[ResultIndex],
    Snapshot := FResultSnapshot)
    AND IsEventUnchanged(Event := FEvents[AggregationIndex],
        Snapshot := FAggregationSnapshot);
END_METHOD

{region 'Documentation'}
(*!
<summary>Initializes the checking Assertions; the scenario explicitly initializes its isolated subject.</summary>
*)
{endregion}
METHOD PROTECTED Configure
FPreparationStateCount := 0;
FTestStateCount := 1;
FLifecycle.Initialize(Parent := THIS^,
    AssertionName := 'Lifecycle');
FPublication.Initialize(Parent := THIS^,
    AssertionName := 'Publication');
FEventOrder.Initialize(Parent := THIS^,
    AssertionName := 'EventOrder');
FFrozenPayload.Initialize(Parent := THIS^,
    AssertionName := 'FrozenPayload');
FStatusRefresh.Initialize(Parent := THIS^,
    AssertionName := 'StatusRefresh');
FChildCalls.Initialize(Parent := THIS^,
    AssertionName := 'ChildCalls');
FCleanup.Initialize(Parent := THIS^,
    AssertionName := 'Cleanup');
END_METHOD

{region 'Documentation'}
(*!
<summary>Compares every defined event field with the retained publication snapshot, without padding or pointer comparisons.</summary>
*)
{endregion}
METHOD PRIVATE IsEventUnchanged : BOOL //! TRUE when all defined event fields match the retained snapshot; structure padding is ignored.
VAR_IN_OUT CONSTANT
    Event : ST_Event; //! Borrowed read-only event to compare field by field.
    Snapshot : ST_Event; //! Borrowed read-only publication snapshot used as the expected value.
END_VAR
IsEventUnchanged := (Event.SequenceId = Snapshot.SequenceId) AND (Event.Timestamp = Snapshot.Timestamp)
    AND (Event.OwnerScope = Snapshot.OwnerScope) AND (Event.EventType = Snapshot.EventType)
    AND (Event.Severity = Snapshot.Severity) AND (Event.Name = Snapshot.Name)
    AND (Event.ResourceName = Snapshot.ResourceName) AND (Event.State = Snapshot.State)
    AND (Event.Result = Snapshot.Result) AND (Event.Message = Snapshot.Message);
END_METHOD

{region 'Documentation'}
(*!
<summary>No asynchronous test resource remains to stop.</summary>
*)
{endregion}
METHOD PROTECTED ProcessAbort
VAR_INPUT
    Enable : BOOL; //! Phase permission supplied by the owning Test Case; FALSE does not authorize progression, while observation may continue.
END_VAR
IF Enable THEN
    CompleteAbort();
END_IF;
END_METHOD

{region 'Documentation'}
(*!
<summary>Checks each observation before advancing; assertions latch across the entire scenario.</summary>
*)
{endregion}
METHOD PROTECTED ProcessAssertions
VAR_INPUT
    Enable : BOOL; //! Phase permission supplied by the owning Test Case; FALSE does not authorize progression, while observation may continue.
END_VAR
FLifecycle(Enable := Enable,
    State := State,
    IN := FLifecycleMatches);
FPublication(Enable := Enable,
    State := State,
    IN := FPublicationMatches);
FEventOrder(Enable := Enable,
    State := State,
    IN := FEventOrderMatches);
FFrozenPayload(Enable := Enable,
    State := State,
    IN := FFrozenPayloadMatches);
FStatusRefresh(Enable := Enable,
    State := State,
    IN := FStatusRefreshMatches);
FChildCalls(Enable := Enable,
    State := State,
    IN := FChildCallsMatches);
FCleanup(Enable := Enable,
    State := State,
    IN := FCleanupMatches);
IF Enable THEN
    FStepChecked := TRUE;
END_IF;
END_METHOD

{region 'Documentation'}
(*!
<summary>No resource Preparation is required for this controlled owner scenario.</summary>
*)
{endregion}
METHOD PROTECTED ProcessPreparations
VAR_INPUT
    // SA0033: Required override; the scenario has no Preparation phase.
    {attribute 'analysis' := '-33'}
    Enable : BOOL; //! Phase permission supplied by the owning Test Case; FALSE does not authorize progression, while observation may continue.
END_VAR
END_METHOD

{region 'Documentation'}
(*!
<summary>Restarts the test script and clears checking Assertions; subject setup belongs to the next test attempt.</summary>
*)
{endregion}
METHOD PROTECTED ProcessReset
FStep := Setup;
FNextStep := Setup;
FStepChecked := FALSE;
FSubjectCalls := 0;
FExpectFinalization := FALSE;
FExpectCompletion := FALSE;
FSavedFinalization := FALSE;
FFinalizationCall := 0;
FCompletedSequence := 0;
FLifecycleMatches := TRUE;
FPublicationMatches := TRUE;
FEventOrderMatches := TRUE;
FFrozenPayloadMatches := TRUE;
FStatusRefreshMatches := TRUE;
FChildCallsMatches := TRUE;
FCleanupMatches := TRUE;
FLifecycle.Reset();
FPublication.Reset();
FEventOrder.Reset();
FFrozenPayload.Reset();
FStatusRefresh.Reset();
FChildCalls.Reset();
FCleanup.Reset();
CompleteReset();
END_METHOD

{region 'Documentation'}
(*!
<summary>Advances the explicit test script with at most one subject FB call per active PLC cycle.</summary>
*)
{endregion}
METHOD PROTECTED ProcessTests
VAR_INPUT
    Enable : BOOL; //! Phase permission supplied by the owning Test Case; FALSE does not authorize progression, while observation may continue.
END_VAR
IF NOT Enable THEN
    RETURN;
END_IF;
IF FStepChecked THEN
    FStep := FNextStep;
    FStepChecked := FALSE;
END_IF;
IF FStep = Done THEN
    CompleteTests();
    RETURN;
END_IF;
RunStep();
END_METHOD

{region 'Documentation'}
(*!
<summary>Runs one subject cycle with fixed expectations; only the Reset-timeout checkpoint may repeat.</summary>
*)
{endregion}
METHOD PRIVATE RunStep
VAR
    Config : ST_TestSuiteConfig;
    Snapshot : ST_TestSuiteStatus;
    ExpectedState : E_State;
    ExpectedResult : E_Result;
    ExpectedTask : E_OrchestratorTask;
    Released : BOOL;
END_VAR
FNextStep := FStep + 1;
ExpectedResult := E_Result.NotEvaluated;
ExpectedTask := E_OrchestratorTask.Idle;

CASE FStep OF
    Setup:
        FExpectedFinalResult := E_Result.Passed;
        IF LateResetChildren THEN
            Config.ResetTimeout := T#50ms;
            FExpectedFinalResult := E_Result.Error;
        END_IF;
        IF NOT FCapture.Initialize(Buffer := FEvents,
            FifoControl := FCaptureFifo,
            Status := FCaptureStatus) THEN
            Error(Message := 'Suite finalization capture could not be initialized.');
            RETURN;
        END_IF;
        FHelper.BeginScenario();
        FSubject.Bind(Publisher := FCapture,
            Helper := FHelper);
        IF NOT FSubject.Initialize(Parent := FSubjectParent,
            SuiteName := 'FinalizationSubject',
            Config := Config) THEN
            Error(Message := 'Suite finalization subject could not be initialized.');
            RETURN;
        END_IF;
        FFirstChild.State := E_State.Uninitialized;
        FFirstChild.Result := E_Result.NotEvaluated;
        FFirstChild.Ready := FALSE;
        FFirstChild.Complete := FALSE;
        FSecondChild := FFirstChild;
        ExpectedState := E_State.Uninitialized;

    ResetRequested:
        IF FSubject.ReserveResetEvents() <> E_EventReservationResult.Accepted THEN
            Error(Message := 'Suite finalization Reset reservation was rejected.');
            RETURN;
        END_IF;
        FSubject.RequestReset();
        FFirstChild.State := E_State.Reset;
        FSecondChild := FFirstChild;
        ExpectedState := E_State.Reset;
        ExpectedTask := E_OrchestratorTask.Reset;

    ResetOutcome:
        IF LateResetChildren THEN
            ExpectedState := E_State.Completing;
            ExpectedResult := E_Result.Error;
            FNextStep := CompleteState;
        ELSE
            FHelper.SetObservation(Ready := TRUE,
                ResetFinished := TRUE);
            FFirstChild.State := E_State.Idle;
            FFirstChild.Ready := TRUE;
            FSecondChild := FFirstChild;
            ExpectedState := E_State.Idle;
        END_IF;

    StartRequested:
        IF FSubject.ReserveExecutionEvents() <> E_EventReservationResult.Accepted THEN
            Error(Message := 'Suite finalization execution reservation was rejected.');
            RETURN;
        END_IF;
        FSubject.RequestStart();
        FFirstChild.State := E_State.Running;
        FFirstChild.Ready := FALSE;
        ExpectedState := E_State.Starting;
        ExpectedTask := E_OrchestratorTask.Execution;

    CompleteChildren:
        FHelper.SetObservation(Ready := FALSE);
        FFirstChild.State := E_State.Completed;
        FFirstChild.Result := E_Result.Passed;
        FFirstChild.Ready := FALSE;
        FFirstChild.Complete := TRUE;
        FSecondChild := FFirstChild;
        ExpectedState := E_State.Running;
        ExpectedTask := E_OrchestratorTask.Execution;

    CompleteOwner:
        FHelper.SetObservation(Ready := FALSE,
            ExecutionFinished := TRUE);
        ExpectedState := E_State.Completing;
        ExpectedResult := E_Result.Passed;
        ExpectedTask := E_OrchestratorTask.Execution;
        FExpectFinalization := TRUE;

    CompleteState:
        ExpectedState := E_State.Completed;
        ExpectedResult := FExpectedFinalResult;
        FExpectCompletion := TRUE;

    LateChildProgress, QuietCompleted, ReleaseReservations, QuietAfterRelease:
        IF LateResetChildren THEN
            FFirstChild.State := E_State.Completed;
            FFirstChild.Result := E_Result.Error;
            FFirstChild.Complete := TRUE;
            FSecondChild.State := E_State.Idle;
            FSecondChild.Ready := TRUE;
        END_IF;
        ExpectedState := E_State.Completed;
        ExpectedResult := FExpectedFinalResult;
ELSE
    Error(Message := 'Unexpected Suite finalization step.');
    RETURN;
END_CASE;

FSubject.SetChildObservations(FirstChild := FFirstChild,
    SecondChild := FSecondChild);
FSubject();
FSubjectCalls := FSubjectCalls + 1;
Snapshot := FSubject.Status;

IF (FStep = ResetOutcome) AND LateResetChildren THEN
    IF FSubject.State = E_State.Reset THEN
        ExpectedState := E_State.Reset;
        ExpectedTask := E_OrchestratorTask.Reset;
        ExpectedResult := E_Result.NotEvaluated;
        FNextStep := ResetOutcome;
    ELSE
        FExpectFinalization := TRUE;
        FLifecycleMatches := FLifecycleMatches AND FSubject.HasResetTimeout;
    END_IF;
END_IF;
FLifecycleMatches := FLifecycleMatches AND (FSubject.State = ExpectedState)
    AND (Snapshot.Execution.State = ExpectedState) AND (FSubject.Result = ExpectedResult)
    AND (FHelper.CurrentTask = ExpectedTask);
FChildCallsMatches := (FSubject.ChildCallCount = FSubjectCalls)
    AND (FHelper.ExecuteCount = FSubjectCalls) AND FSubject.ChildBodyCallsMatch;

IF FExpectFinalization AND NOT FSavedFinalization THEN
    IF LateResetChildren THEN
        FExpectedAggregation := '{"total":2,"inactive":0,"idle":0,"running":0,"completed":0,"passed":0,"failed":0,"error":0,"runtime":';
    ELSE
        FExpectedAggregation := '{"total":2,"inactive":0,"idle":0,"running":0,"completed":2,"passed":2,"failed":0,"error":0,"runtime":';
    END_IF;
    FExpectedAggregation := CONCAT(FExpectedAggregation, UDINT_TO_STRING(TIME_TO_UDINT(Snapshot.Runtime)));
    FExpectedAggregation := CONCAT(FExpectedAggregation, '}');
END_IF;
CheckEventStream();

